(* IEC 61131-3 sources: plcassist-cli/packages/volt-lsp-iec/test-corpus/awa-palletizer/Device/Plc Logic/Application/Library Manager/AlarmManager (part 3) *)

(* ---- DATABASEFILEALARMSTORAGE.fb ---- *)
FUNCTION_BLOCK DATABASEFILEALARMSTORAGE EXTENDS AlarmStorageManager
VAR
	M_SAPPLICATIONNAME : STRING;
	M_AITFALARMSTORAGELISTENER : ARRAY [0..(COUNT_MAX_ALARM_STORAGE_LISTENER - 1)] OF IAlarmStorageListener;
	M_SOLDREMOTEDEVICENAME : STRING;
	M_LIREMOTEDEVICENAMEVALUE : LINT;
	M_CACHEDDBVERSION : INT := UNDETERMINED_DB_VERSION;
	M_CACHEDDBVERSIONERROR : STO.ERROR;
	M_WRITECONTEXT : DatabaseFileWriteContext;
	M_XCHANGESTATETONORMAL : BOOL;
	M_XASSIGNINACTIVETIMESTAMPS : BOOL;
	COUNT_MAX_ALARM_STORAGE_LISTENER : INT := 5;
	UNDETERMINED_DB_VERSION : INT := -1;
	ASSIGNINACTIVETIMESTAMPS : BOOL;
	CHANGESTATETONORMAL : BOOL;
	TABLE : STO.ITable;
	WRITEACCESSNECESSARY : BOOL;
END_VAR
END_FUNCTION_BLOCK

METHOD GETDATABASEFILEPATH : STRING
END_METHOD

METHOD GETFILELIMIT : FileLimit
END_METHOD

METHOD GETMAXRECORDCOUNT : UDINT
END_METHOD

METHOD GETSUBDIRECTORY : STRING
END_METHOD

METHOD WRITETOSTORAGE : STO.ERROR
VAR_INPUT
	ITFTABLE : STO.ITable;
	ROW : AlarmStorageRow;
	ICOUNTRETRIES : INT;
END_VAR
END_METHOD

METHOD CLEARBUFFER
END_METHOD

METHOD ADDALARMSTORAGELISTENER : EAlarmStorageReaderErrors
VAR_INPUT
	ITFALARMSTORAGELISTENER : IAlarmStorageListener;
END_VAR
END_METHOD

METHOD CREATEALARMSTORAGEMETADATAFILE
VAR_INPUT
	UDICOUNTCOLUMNSTBLALARM : CAA.COUNT;
END_VAR
END_METHOD

METHOD OPENTABLE2 : STO.ITable
VAR_INPUT
	XREADONLY : BOOL;
END_VAR
VAR_OUTPUT
	EERROR : STO.ERROR;
END_VAR
END_METHOD

METHOD REMOVEALARMSTORAGELISTENER : EAlarmStorageReaderErrors
VAR_INPUT
	ITFALARMSTORAGELISTENER : IAlarmStorageListener;
END_VAR
END_METHOD

METHOD CHECKFILELIMITREACHED : STO.Error
VAR_INPUT
	ITFTABLE : STO.ITable;
	ICOUNTRETRIES : INT;
	ICOUNTROWSTOINSERT : INT;
END_VAR
END_METHOD

METHOD GETEXCLUSIVETRANSACTION : STO.ITransaction
VAR_INPUT
	ICOUNTRETRIES : INT;
END_VAR
VAR_OUTPUT
	EERROR : STO.ERROR;
END_VAR
END_METHOD

METHOD WRITETOSTORAGE2 : STO.ERROR
VAR_INPUT
	ITFTABLE : STO.ITable;
	ROW : AlarmStorageRow;
	ITFTRANSACTION : STO.ITransaction;
END_VAR
END_METHOD

METHOD DELETEALARMSTORAGEFILE : STO.ERROR
VAR_INPUT
	SFILEPATH : CAA.FILENAME;
END_VAR
END_METHOD

METHOD GETALARMSFROMSTORAGE : STO.ERROR
VAR_INPUT
	ISKIPROWS : INT;
	IMAXROWS : INT;
	FILTERCRITERIA : REFERENCE TO VisuFbAlarmFilterCriteria;
	ITFALARMDATABLOCK : IAlarmDataBlockBase2;
END_VAR
VAR_IN_OUT
	BROWIDVALID : BOOL;
	DIROWID : DINT;
END_VAR
END_METHOD

METHOD GETCOUNTALARMSFROMSTORAGE : DINT
VAR_INPUT
	FILTERCRITERIA : REFERENCE TO VisuFbAlarmFilterCriteria;
	ITFALARMDATABLOCK : IAlarmDataBlockBase2;
END_VAR
VAR_OUTPUT
	EERROR : STO.ERROR;
	DWCOUNTLATCHVARIABLESINSTORAGE : CAA.COUNT;
END_VAR
END_METHOD

METHOD CREATEWRITECONTEXT : IDatabaseFileWriteContext
END_METHOD

METHOD SCANSTORAGE : STO.ERROR
VAR_INPUT
	ITFCONSUMER : IRemoteDeviceTraversalConsumer;
END_VAR
VAR_OUTPUT
	IVERSION : INT;
	DIREMOTEENTRIESCNT : DINT;
END_VAR
END_METHOD

METHOD WRITETOSTORAGE3 : STO.ERROR
VAR_INPUT
	WRITECONTEXT : IDatabaseFileWriteContext;
	ROW : AlarmStorageRow;
	XFORCEINSERT : BOOL;
	XFIRST : BOOL;
END_VAR
END_METHOD

METHOD CLEARALARMSINSTATENORMAL : STO.Error
VAR_INPUT
	ITFTABLE : STO.ITable;
END_VAR
VAR_OUTPUT
	XFINISHED : BOOL;
END_VAR
VAR_IN_OUT
	DIREMAININGROWCOUNT : DINT;
END_VAR
END_METHOD

METHOD ROWSELECT : STO.IRow
VAR_INPUT
	ITFTABLE : STO.ITable;
	IDROW : CAA.IDENT;
END_VAR
END_METHOD

METHOD CHECKRECORDLIMITREACHED : STO.Error
VAR_INPUT
	ITFTABLE : STO.ITable;
	ICOUNTRETRIES : INT;
	ICOUNTROWSTOINSERT : INT;
	XFORCE : BOOL;
END_VAR
VAR_OUTPUT
	XLIMIT : BOOL;
	UDIMAXRECORDCOUNT : UDINT;
END_VAR
END_METHOD

METHOD DELETEALARMS : STO.Error
VAR_INPUT
	ITFTABLE : STO.ITable;
	ICOUNTRETRIES : INT;
	DICOUNTROWSTODELETE : DINT;
END_VAR
VAR_OUTPUT
	DIROWSDELETED : DINT;
END_VAR
END_METHOD

METHOD GETRECORDSIZE : INT
END_METHOD

METHOD GETSTORAGESIZE : LINT
END_METHOD

METHOD SETEMPTYTIMESTAMPINACTIVETOSTARTTIME : STO.Error
VAR_INPUT
	ITFTABLE : STO.ITable;
END_VAR
END_METHOD

METHOD CHECKFILELIMITREACHEDUDINT : STO.ERROR
VAR_INPUT
	ITFTABLE : STO.ITable;
	ICOUNTRETRIES : INT;
	UDICOUNTROWSTOINSERT : UDINT;
END_VAR
END_METHOD

METHOD CHECKRECORDLIMITREACHEDUDINT : STO.ERROR
VAR_INPUT
	ITFTABLE : STO.ITable;
	ICOUNTRETRIES : INT;
	UDICOUNTROWSTOINSERT : UDINT;
	XFORCE : BOOL;
END_VAR
VAR_OUTPUT
	XLIMIT : BOOL;
	UDIMAXRECORDCOUNT : UDINT;
END_VAR
END_METHOD

METHOD PRVCHECKFILELIMITREACHED : STO.Error
VAR_INPUT
	ITFTABLE : STO.ITable;
	ICOUNTRETRIES : INT;
	UDICOUNTROWSTOINSERT : UDINT;
END_VAR
END_METHOD

METHOD PRVCHECKRECORDLIMITREACHED : STO.Error
VAR_INPUT
	ITFTABLE : STO.ITable;
	ICOUNTRETRIES : INT;
	UDICOUNTROWSTOINSERT : UDINT;
	XFORCE : BOOL;
END_VAR
VAR_OUTPUT
	XLIMIT : BOOL;
	UDIMAXRECORDCOUNT : UDINT;
END_VAR
END_METHOD

METHOD PRVDELETEALARMSTOREACHLIMIT : BOOL
VAR_INPUT
	ITFTABLE : STO.ITable;
	ICOUNTRETRIES : INT;
	UDICOUNTROWSTODELETE : UDINT;
END_VAR
VAR_OUTPUT
	IROWSDELETED : INT;
	EERROR : STO.ERROR;
END_VAR
END_METHOD

METHOD PRVFINDLATCHVARSTRING
VAR_INPUT
	CBPINPUTSTRING : CharBufferPtr;
	BYTYPECLASS : BYTE;
	IVERSION : INT;
	ITFTABLE : STO.ITable;
END_VAR
VAR_OUTPUT
	DIROWID : DINT;
	XFOUND : BOOL;
END_VAR
VAR_IN_OUT
	EERROR : STO.ERROR;
	WSINPUTSTRING : WSTRING(255);
END_VAR
END_METHOD

METHOD PRVFINDLATCHVARSTRING_DBVERBEFORE5
VAR_INPUT
	CBPINPUTSTRING : CharBufferPtr;
	BYTYPECLASS : BYTE;
	ITFCURSOR : STO.ICursor;
END_VAR
VAR_OUTPUT
	DIROWID : DINT;
	XFOUND : BOOL;
END_VAR
VAR_IN_OUT
	EERROR : STO.ERROR;
END_VAR
END_METHOD

METHOD PRVFINDLATCHVARSTRING_DBVERRECENT
VAR_INPUT
	ITFCURSOR : STO.ICursor;
END_VAR
VAR_OUTPUT
	DIROWID : DINT;
	XFOUND : BOOL;
END_VAR
VAR_IN_OUT
	EERROR : STO.ERROR;
	WSINPUTSTRING : WSTRING(255);
END_VAR
END_METHOD

METHOD PRVGETDATABASEFILEPATH : STRING
VAR_INPUT
	SVERSIONINCOMPATIBLECHANGE : STRING;
END_VAR
VAR_OUTPUT
	EERROR : STO.ERROR;
END_VAR
END_METHOD

METHOD PRVGETVERSION : STO.ERROR
VAR_OUTPUT
	IVERSION : INT;
END_VAR
END_METHOD

METHOD PRVGETVERSIONFROMDATABASE : STO.ERROR
VAR_OUTPUT
	IVERSION : INT;
END_VAR
END_METHOD

METHOD PRVREMOVERECORDLIMITREACHED : STO.Error
VAR_INPUT
	UDIMAXRECORDCOUNT : UDINT;
	ITFTABLE : STO.ITable;
	ICOUNTRETRIES : INT;
	ICOUNTROWSTOINSERT : UDINT;
END_VAR
END_METHOD

METHOD PRVSEARCHMINROWIDS : STO.ERROR
VAR_INPUT
	ITFTABLE : STO.ITable;
	ICOUNTROWSIDSTOSEARCH : INT;
	PADWROWIDS : POINTER TO ARRAY [0..50] OF CAA.IDENT;
	IEFFECTIVEARRAYSIZE : INT;
END_VAR
VAR_OUTPUT
	ICOUNTROWSIDS : INT;
END_VAR
END_METHOD

METHOD PRVSETTYPEDVALUE : STO.ERROR
VAR_INPUT
	BYTYPECLASS : BYTE;
	LIVALUE : LINT;
	ITFROWBASE : STO.IRowBase;
	COLVALUE : CAA.IDENT;
	COLTYPE : CAA.IDENT;
END_VAR
END_METHOD

METHOD PRVSORTROWIDS
VAR_INPUT
	PADWROWIDS : POINTER TO ARRAY [0..0] OF CAA.IDENT;
	NFIRST : INT;
	NLAST : INT;
END_VAR
END_METHOD

METHOD PRVSTOREALARMCOMMENTS : STO.ERROR
VAR_INPUT
	PROW : POINTER TO AlarmStorageRow;
	ITFROWPLANCHET : STO.IRowPlanchet;
	ITFROW : STO.IRow;
END_VAR
END_METHOD

METHOD PRVUPDATEROW : BOOL
VAR_INPUT
	HTASK : RTS_IEC_HANDLE;
	ITFROW : STO.IRow;
	ICOUNTRETRIES : INT;
	EERROR : STO.ERROR;
END_VAR
END_METHOD

METHOD PRVWRITEALARMCOMMENTCOLUMN
VAR_INPUT
	PWSVALUE : POINTER TO WSTRING;
	ITFROWPLANCHET : STO.IRowPlanchet;
	ITFROW : STO.IRow;
	DATABASEIDENT : CAA.IDENT;
	ERRACTION : INT;
END_VAR
VAR_IN_OUT
	EERROR : STO.ERROR;
END_VAR
END_METHOD

METHOD PRVWRITEBYTEORDERFLAG
END_METHOD

METHOD PRVWRITELATCHVARSTRINGS
VAR_INPUT
	ITFROWBASE : STO.IRowBase;
	PROW : POINTER TO AlarmStorageRow;
	WRITECONTEXT : IDatabaseFileWriteContext;
END_VAR
VAR_IN_OUT
	EERROR : STO.ERROR;
END_VAR
END_METHOD

METHOD PRVWRITETOSTORAGE : STO.ERROR
VAR_INPUT
	WRITECONTEXT : IDatabaseFileWriteContext;
	ROW : AlarmStorageRow;
	ICOUNTRETRIES : INT;
	XCHECKFILELIMITREACHED : BOOL;
	XFORCEINSERT : BOOL;
END_VAR
END_METHOD

METHOD PRVWRITETOTBLLATCHVARSTRINGS : STO.ERROR
VAR_INPUT
	WRITECONTEXT : IDatabaseFileWriteContext;
	CBPINPUTSTRING : CharBufferPtr;
	BYTYPECLASS : BYTE;
END_VAR
VAR_OUTPUT
	DIROWID : DINT;
END_VAR
END_METHOD

METHOD PRVWRITETRIGGERVALUE
VAR_INPUT
	ITFROWBASE : STO.IRowBase;
	BYTRIGGERVALUETYPE : BYTE;
	LITRIGGERVALUEVAL : LINT;
END_VAR
VAR_IN_OUT
	EERROR : STO.ERROR;
END_VAR
END_METHOD

(* ---- DATABASEFILEWRITECONTEXT.fb ---- *)
FUNCTION_BLOCK DATABASEFILEWRITECONTEXT EXTENDS DatabaseFileWriteContextBase
VAR
	_INUSE : BOOL;
	M_ICOUNTRETRIES : INT := AlarmConstants.RETRY_COUNT;
	M_ICOUNTCYCLEWAIT : INT;
END_VAR
END_FUNCTION_BLOCK

METHOD INITIALIZE : BOOL
VAR_IN_OUT
	DB : DatabaseFileAlarmStorage;
END_VAR
END_METHOD

METHOD RELEASE
VAR_INPUT
	EERRORFORCOMMIT : STO.ERROR;
END_VAR
END_METHOD

METHOD PRVINCREASERETRYCOUNT : BOOL
END_METHOD

METHOD PRVRESETRETRYCOUNT : BOOL
END_METHOD

(* ---- DATABASEFILEWRITECONTEXTBASE.fb ---- *)
FUNCTION_BLOCK DATABASEFILEWRITECONTEXTBASE
VAR
	_MAINTABLE : STO.ITable;
	_STRINGLATCHTABLE : STO.ITable;
	_TRANSACTION : STO.ITransaction;
	_STORAGEMAN : REFERENCE TO DatabaseFileAlarmStorage;
	MAINTABLE : STO.ITable;
	TRANSACTION : STO.ITransaction;
END_VAR
END_FUNCTION_BLOCK

METHOD GETSTRINGLATCHTABLE : STO.ITable
VAR_OUTPUT
	EERROR : STO.ERROR;
END_VAR
END_METHOD

METHOD RELEASE
VAR_INPUT
	EERRORFORCOMMIT : STO.ERROR;
END_VAR
END_METHOD

(* ---- DATABASEFILEWRITECONTEXTTEMPORARY.fb ---- *)
FUNCTION_BLOCK DATABASEFILEWRITECONTEXTTEMPORARY EXTENDS DatabaseFileWriteContextBase
END_FUNCTION_BLOCK

METHOD FB_EXIT : BOOL
VAR_INPUT
	BINCOPYCODE : BOOL;
END_VAR
END_METHOD

METHOD INITIALIZE : BOOL
VAR_INPUT
	MAINTABLE : STO.ITable;
	TRANSACTION : STO.ITransaction;
END_VAR
VAR_IN_OUT
	STORAGEMAN : DatabaseFileAlarmStorage;
END_VAR
END_METHOD

(* ---- DATABASESIZELIMIT.fb ---- *)
FUNCTION_BLOCK DATABASESIZELIMIT
VAR
	M_XINITIALIZED : BOOL;
	M_XFIRST : BOOL := TRUE;
	M_XFIRSTREMOVE : BOOL := TRUE;
	M_METRICS : STO.METRICS;
	M_ITFDATABASEFILEALARMSTORAGE7 : IDatabaseFileAlarmStorage7;
	M_ITFALARMSTORAGEMANAGER : IAlarmStorageManager;
	M_SYSRECORDSIZE : INT;
	M_LISTORAGESIZE : LINT;
	M_XERRORDISPLAYED : BOOL;
	M_LIFILESIZEINERROR : LINT;
	M_ICNTREORGERR : INT;
	M_XBLOCKED : BOOL;
	M_ITEMPREDUCTIONRECORDNUM : INT;
	M_TLASTREORGTIME : TIME;
	M_ICNTDBREORD : INT;
	ISBLOCKED : BOOL;
	LASTREORDERINGTIME : TIME;
	REORDERINGCOUNT : INT;
END_VAR
END_FUNCTION_BLOCK

METHOD CHECKFORSIZELIMIT : BOOL
END_METHOD

METHOD INITIALIZE
VAR_INPUT
	ITFDATABASEFILEALARMSTORAGE : IDatabaseFileAlarmStorage;
END_VAR
END_METHOD

METHOD PRVDBMETRICS : STO.ERROR
VAR_OUTPUT
	MMETRICS : STO.METRICS;
END_VAR
END_METHOD

METHOD PRVGETRECORDSIZE : INT
END_METHOD

METHOD PRVGETRECORDSTOREMOVE : DINT
VAR_INPUT
	LIBYTESTOREMOVE : LINT;
END_VAR
VAR_OUTPUT
	IRECORDSIZE : INT;
END_VAR
END_METHOD

METHOD PRVREORGDB : STO.ERROR
END_METHOD

(* ---- DEFAULTALARMFILTERCRITERIA.fb ---- *)
FUNCTION_BLOCK DEFAULTALARMFILTERCRITERIA
END_FUNCTION_BLOCK

METHOD AREALLALARMCLASSESSELECTED : BOOL
END_METHOD

METHOD AREALLALARMGROUPSSELECTED : BOOL
END_METHOD

METHOD GETALARMCLASSES : POINTER TO ARRAY [0..0] OF UDINT
END_METHOD

METHOD GETALARMGROUPS : POINTER TO ARRAY [0..0] OF UDINT
END_METHOD

METHOD GETCOUNTALARMCLASSES : INT
END_METHOD

METHOD GETCOUNTALARMGROUPS : INT
END_METHOD

METHOD GETPRIORITYFROM : USINT
END_METHOD

METHOD GETPRIORITYTO : USINT
END_METHOD

(* ---- EVENTDISPATCHER.fb ---- *)
FUNCTION_BLOCK EVENTDISPATCHER
VAR
	_HGETCOUNTEVENT : RTS_IEC_HANDLE := Events.Invalid_Handle;
	_HGETCOUNTEVENTINTERFACE : RTS_IEC_HANDLE := Events.Invalid_Handle;
	_HGETALARMSEVENT : RTS_IEC_HANDLE := Events.Invalid_Handle;
	_HGETALARMSEVENTINTERFACE : RTS_IEC_HANDLE := Events.Invalid_Handle;
	_HCHANNELCLOSEDEVENT : RTS_IEC_HANDLE := Events.Invalid_Handle;
	_HCHANNELCLOSEDEVENTINTERFACE : RTS_IEC_HANDLE := Events.Invalid_Handle;
	_HHANDLESERVICEEVENT : RTS_IEC_HANDLE := Events.Invalid_Handle;
	_HHANDLESERVICEEVENTINTERFACE : RTS_IEC_HANDLE := Events.Invalid_Handle;
	_SERVICEHANDLER : AlarmServiceHandler;
END_VAR
END_FUNCTION_BLOCK

METHOD EVENTCALLBACK : UDINT
VAR_INPUT
	PEVENTPARAM : POINTER TO EventParam;
END_VAR
END_METHOD

METHOD FB_EXIT : BOOL
VAR_INPUT
	BINCOPYCODE : BOOL;
END_VAR
END_METHOD

METHOD FB_INIT : BOOL
VAR_INPUT
	BINITRETAINS : BOOL;
	BINCOPYCODE : BOOL;
END_VAR
END_METHOD

(* ---- EXPRESSIONOBSERVATIONTYPE.fb ---- *)
FUNCTION_BLOCK EXPRESSIONOBSERVATIONTYPE
VAR_INPUT
	M_UIID : ALARM_ID;
	M_EXPRESSIONEVALUATOR : IExpressionEvaluator;
END_VAR
END_FUNCTION_BLOCK

METHOD ISACTIVE : BOOL
VAR_INPUT
	ECURRSTATE : AlarmState;
END_VAR
END_METHOD

METHOD ISIMMEDIATELYACTIVE : BOOL
END_METHOD

(* ---- FORMATSTRINGSCANNER.fb ---- *)
FUNCTION_BLOCK FORMATSTRINGSCANNER
END_FUNCTION_BLOCK

METHOD GETFORMATSTRING : BOOL
VAR_INPUT
	RCBSMESSAGE : REFERENCE TO CharBufferString;
	PCBSPLACEHOLDER : POINTER TO CharBufferString;
	IOFFSET : INT;
	ILENGTHPREFIX : INT;
END_VAR
VAR_OUTPUT
	SFORMATSTRING : STRING;
	ITOTALPLACEHOLDERLENGTH : INT;
END_VAR
END_METHOD

(* ---- HASHTABLEKEYELEMENT.fb ---- *)
FUNCTION_BLOCK HASHTABLEKEYELEMENT EXTENDS InstanceBase
VAR
	_INSTANCEPOINTER : POINTER TO BYTE;
	_ALARMTEMPLATENAME : POINTER TO STRING;
	_LIHASH : LINT;
	ALARMTEMPLATENAME : POINTER TO STRING;
	INSTANCEPOINTER : POINTER TO BYTE;
END_VAR
END_FUNCTION_BLOCK

METHOD ELEMENTCOMPARETO : INT
VAR_INPUT
	ITFELEMENT : COL.IElement;
END_VAR
END_METHOD

METHOD ELEMENTEQUALS : BOOL
VAR_INPUT
	ITFELEMENT : COL.IElement;
END_VAR
END_METHOD

METHOD ELEMENTHASHCODE : LINT
END_METHOD

METHOD PRVCALCULATEHASH : LINT
END_METHOD

METHOD PRVINSTINIT : COL.FBF.ERROR
VAR_INPUT
	ITFDATA : COL.FBF.IData;
END_VAR
END_METHOD

(* ---- HASHTABLEKEYELEMENTDATA.fb ---- *)
FUNCTION_BLOCK HASHTABLEKEYELEMENTDATA EXTENDS InstanceData
VAR_INPUT
	PALARMINSTANCE : POINTER TO BYTE;
	STALARMTEMPLATENAME : POINTER TO STRING;
END_VAR
END_FUNCTION_BLOCK

(* ---- HASHTABLEKEYELEMENTFACTORY.fb ---- *)
FUNCTION_BLOCK HASHTABLEKEYELEMENTFACTORY EXTENDS FactoryBase
VAR
	PRVINSTCOUNT : CAA.COUNT;
	PRVINSTPOOLEXTENDSFACTOR : USINT;
	PRVINSTSIZE : CAA.SIZE;
END_VAR
END_FUNCTION_BLOCK

METHOD CREATE : IHashtableKeyElement
VAR_INPUT
	INSTANCEPOINTER : POINTER TO BYTE;
	PSTALARMTEMPLATENAME : POINTER TO STRING;
END_VAR
VAR_OUTPUT
	EERROR : COL.FBF.ERROR;
END_VAR
END_METHOD

(* ---- HASHTABLEVALUEELEMENT.fb ---- *)
FUNCTION_BLOCK HASHTABLEVALUEELEMENT EXTENDS InstanceBase
VAR
	_UDIALARMGROUPID : UDINT;
	_UITEMPLATEALARMSOFFSET : UINT;
	_UITEMPLATEALARMSLENGTH : UINT;
	_UITEMPLATEEVENTSOFFSET : UINT;
	_UITEMPLATEEVENTSLENGTH : UINT;
	ALARMGROUPID : UDINT;
	TEMPLATEALARMSLENGTH : UINT;
	TEMPLATEALARMSOFFSET : UINT;
	TEMPLATEEVENTSLENGTH : UINT;
	TEMPLATEEVENTSOFFSET : UINT;
END_VAR
END_FUNCTION_BLOCK

METHOD ELEMENTCOMPARETO : INT
VAR_INPUT
	ITFELEMENT : COL.IElement;
END_VAR
END_METHOD

METHOD ELEMENTEQUALS : BOOL
VAR_INPUT
	ITFELEMENT : COL.IElement;
END_VAR
END_METHOD

METHOD ELEMENTHASHCODE : LINT
END_METHOD

METHOD PRVINSTINIT : COL.FBF.ERROR
VAR_INPUT
	ITFDATA : COL.FBF.IData;
END_VAR
END_METHOD

(* ---- HASHTABLEVALUEELEMENTDATA.fb ---- *)
FUNCTION_BLOCK HASHTABLEVALUEELEMENTDATA EXTENDS InstanceData
VAR_INPUT
	UDIALARMGROUPID : UDINT;
	UITEMPLATEALARMSOFFSET : UINT;
	UITEMPLATEALARMSLENGTH : UINT;
	UITEMPLATEEVENTSOFFSET : UINT;
	UITEMPLATEEVENTSLENGTH : UINT;
END_VAR
END_FUNCTION_BLOCK

(* ---- HASHTABLEVALUEELEMENTFACTORY.fb ---- *)
FUNCTION_BLOCK HASHTABLEVALUEELEMENTFACTORY EXTENDS FactoryBase
VAR
	PRVINSTCOUNT : CAA.COUNT;
	PRVINSTPOOLEXTENDSFACTOR : USINT;
	PRVINSTSIZE : CAA.SIZE;
END_VAR
END_FUNCTION_BLOCK

METHOD CREATE : IHashtableValueElement
VAR_INPUT
	UDIALARMGROUPID : UDINT;
	UITEMPLATEALARMSOFFSET : UINT;
	UITEMPLATEALARMSLENGTH : UINT;
	UITEMPLATEEVENTSOFFSET : UINT;
	UITEMPLATEEVENTSLENGTH : UINT;
END_VAR
VAR_OUTPUT
	EERROR : COL.FBF.ERROR;
END_VAR
END_METHOD

(* ---- HISTORICALALARMMOCK.fb ---- *)
FUNCTION_BLOCK HISTORICALALARMMOCK EXTENDS ProxyFbAlarmHistorical
VAR_INPUT
	M_BALARMSTORAGE : BYTE;
	M_DWROWIDFIRST : DWORD;
	M_DWROWIDLAST : DWORD;
	M_SVALUE : STRING;
	M_WSVALUE : WSTRING;
END_VAR
END_FUNCTION_BLOCK

METHOD SETVALUES
VAR_INPUT
	ISET : INT;
END_VAR
END_METHOD

(* ---- LISTELEMENT.fb ---- *)
FUNCTION_BLOCK LISTELEMENT EXTENDS InstanceBase
VAR
	_ALARMINST : Alarm;
	_USICOUNTLATCHVARIABLES : USINT;
	_ARRLATCHVARIABLES : ARRAY [0..255] OF ValueTypeBundle;
	_XISACTIVEALARM : BOOL;
	ALARM : POINTER TO Alarm;
	ISACTIVEALARM : BOOL;
	ISDEACTIVATEDPREV : BOOL;
END_VAR
END_FUNCTION_BLOCK

METHOD ELEMENTCOMPARETO : INT
VAR_INPUT
	ITFELEMENT : COL.IElement;
END_VAR
END_METHOD

METHOD ELEMENTEQUALS : BOOL
VAR_INPUT
	ITFELEMENT : COL.IElement;
END_VAR
END_METHOD

METHOD ELEMENTHASHCODE : LINT
END_METHOD

METHOD GETLATCHVARIABLES : BOOL
VAR_OUTPUT
	PALATCHVARIABLES : POINTER TO ARRAY [0..255] OF ValueTypeBundle;
	USICOUNTLATCHVARIABLES : USINT;
END_VAR
END_METHOD

METHOD SETLATCHVARIABLES : BOOL
VAR_INPUT
	PALARM : POINTER TO Alarm;
END_VAR
END_METHOD

METHOD PRVINSTINIT : COL.FBF.ERROR
VAR_INPUT
	ITFDATA : COL.FBF.IData;
END_VAR
END_METHOD

(* ---- LISTELEMENTDATA.fb ---- *)
FUNCTION_BLOCK LISTELEMENTDATA EXTENDS InstanceData
END_FUNCTION_BLOCK

(* ---- LISTELEMENTFACTORY.fb ---- *)
FUNCTION_BLOCK LISTELEMENTFACTORY EXTENDS FactoryBase
VAR
	PRVINSTCOUNT : CAA.COUNT;
	PRVINSTPOOLEXTENDSFACTOR : USINT;
	PRVINSTSIZE : CAA.SIZE;
END_VAR
END_FUNCTION_BLOCK

METHOD CREATE : IListElement
VAR_OUTPUT
	EERROR : COL.FBF.ERROR;
END_VAR
END_METHOD

(* ---- MESSAGECOMPARER.fb ---- *)
FUNCTION_BLOCK MESSAGECOMPARER EXTENDS TSLastComparer
VAR
	M_STRINGTYPE : __SYSTEM.TYPE_CLASS;
	M_IWHICHMESSAGE : INT;
	M_ICOUNTLATCHVARIABLES : INT;
	M_CBSMESSAGE1 : CharBufferString;
	M_CBSMESSAGE2 : CharBufferString;
	M_CBSMESSAGE1REPLACED : CharBufferString;
	M_CBSMESSAGE2REPLACED : CharBufferString;
	M_ABYBUFFERMESSAGE1REPLACED : ARRAY [0..(BUFFER_LENGTH - 1)] OF BYTE;
	M_ABYBUFFERMESSAGE2REPLACED : ARRAY [0..(BUFFER_LENGTH - 1)] OF BYTE;
	M_TIMESTAMPANDVALUESCONTAINER : TimestampAndValuesContainer;
	BUFFER_LENGTH : INT := (2 * (255 + 1));
END_VAR
END_FUNCTION_BLOCK

METHOD BEFORECOMPARE
VAR_INPUT
	STRINGTYPE : __SYSTEM.TYPE_CLASS;
	IWHICHMESSAGE : INT;
	ICOUNTLATCHVARIABLES : INT;
END_VAR
END_METHOD

METHOD COMPARE : INT
VAR_INPUT
	DIINDEXALARM1 : DINT;
	DIINDEXALARM2 : DINT;
END_VAR
END_METHOD

METHOD PRVGETALARMMESSAGE : CharBufferPtr
VAR_INPUT
	UDIALARMGROUPID : UDINT;
	UDIALARMID : UDINT;
	SDEVICENAME : STRING;
END_VAR
VAR_OUTPUT
	SALARMID : STRING;
END_VAR
END_METHOD

METHOD PRVREPLACEPLACEHOLDERS : BOOL
VAR_INPUT
	DIINDEXALARM : DINT;
	CBPMESSAGE : CharBufferPtr;
	RCBSMESSAGE : REFERENCE TO CharBufferString;
	RCBSMESSAGEREPLACED : REFERENCE TO CharBufferString;
END_VAR
END_METHOD

(* ---- ONLYDATEANDTIMEPLACEHOLDER.fb ---- *)
FUNCTION_BLOCK ONLYDATEANDTIMEPLACEHOLDER
VAR
	M_APLACEHOLDEROCCURRENCE : ARRAY [PLACEHOLDER_DATE..PLACEHOLDER_TIME] OF PlaceholderOccurrence;
	PLACEHOLDER_DATE : INT := 0;
	PLACEHOLDER_TIME : INT := 1;
END_VAR
END_FUNCTION_BLOCK

METHOD FB_INIT : BOOL
VAR_INPUT
	BINITRETAINS : BOOL;
	BINCOPYCODE : BOOL;
END_VAR
END_METHOD

METHOD ANALYZEPLACEHOLDERS
VAR_INPUT
	STRINGTYPE : __SYSTEM.TYPE_CLASS;
END_VAR
END_METHOD

METHOD GETCOUNTPLACEHOLDERS : SINT
END_METHOD

METHOD GETPLACEHOLDER : PlaceholderOccurrence
VAR_INPUT
	SIWHICHPLACEHOLDER : SINT;
END_VAR
END_METHOD

METHOD HASPLACEHOLDERREQUIRINGCYCLICALLYUPDATE : BOOL
END_METHOD

METHOD HASPLACEHOLDERS : BOOL
END_METHOD

METHOD ISOPTIMIZEDPLACEHOLDERREPLACEMENTSUPPORTED : BOOL
END_METHOD

(* ---- PRIORITYCOMPARER.fb ---- *)
FUNCTION_BLOCK PRIORITYCOMPARER EXTENDS TSLastComparer
END_FUNCTION_BLOCK

METHOD COMPARE : INT
VAR_INPUT
	DIINDEXALARM1 : DINT;
	DIINDEXALARM2 : DINT;
END_VAR
END_METHOD

(* ---- PROXY.fb ---- *)
FUNCTION_BLOCK PROXY
VAR
	M_XISINIT : BOOL;
	M_IRUNSTATUS : INT;
	M_ITFCOMMCHANNEL : IProxyCommChannel;
	M_ITEST : INT;
	M_ESTATE : ProxyEnumState;
	M_SDEVICENAME : STRING;
	M_LIBVERALMMAN : VERSION;
	M_LTSTARTTIMECHANNEL : LTIME;
	M_LTSTARTTIMERUN : LTIME;
	M_LTSTARTTIME : LTIME;
	M_ISTATE : INT;
	M_XALREADYDISP : BOOL;
	M_TTIMEOUT : TIME;
	M_IREQIDSENT : INT;
	M_IREQIDREC : INT;
	M_XWITHERRORS : BOOL;
	M_DWBASETIME : DWORD := (50 * 1000);
	M_DWACTALMTIME : DWORD := (200 * 1000);
	M_DWHISALMTIME : DWORD := (1000 * 1000);
	M_DWACKALMTIME : DWORD := (1000 * 1000);
	M_TGENTIMEOUT : TIME := DEFAULT_TIMEOUT;
	M_APROXYRUNTASKCALL : ARRAY [1..ProxyConstants.MAX_TASK] OF ProxyStructTaskCall;
	M_IRUNTASKCALLMAX : INT;
	M_APROXYPRERUNTASKCALL : ARRAY [1..ProxyConstants.MAX_TASK] OF ProxyStructTaskCall;
	M_IPRERUNTASKCALLMAX : INT;
	M_ITASKCALL : INT;
	M_SPROXYNAME : STRING;
	M_PSAPPNAME : POINTER TO STRING;
	M_CBSMESSAGE : CharBufferString;
	M_AWLOCALBUFFER : ARRAY [0..(LOCAL_TEXT_BUFFER_LENGTH / 2)] OF WORD;
	M_ARECORDS : ARRAY [0..(MAX_RECORDS - 1)] OF ProxyStructRecord;
	M_IRECINUSE : INT;
	M_SIHASSTORAGE : SINT := -1;
	M_DWROWIDFIRSTREMDB : DWORD := AlarmConstants.INVALID_ROWID;
	M_DWROWIDLASTREMDB : DWORD := AlarmConstants.INVALID_ROWID;
	M_DWROWIDLASTVALIDREAD : DWORD := AlarmConstants.INVALID_ROWID;
	M_DWROWIDLASTLOCDB : DWORD := AlarmConstants.INVALID_ROWID;
	M_IROWCOUNTTOREAD : INT;
	M_PAHISTALARMGROUPS : ARRAY [1..MAX_HIST_GROUPS] OF POINTER TO STRING;
	M_IHISTALARMGROUPSNUM : INT;
	M_IHISTRECORDID : INT := -1;
	M_XFIRSTHISTREADDONE : BOOL;
	M_XFIRSTHISTACTIVEREADDONE : BOOL;
	M_XDISP1DONE : BOOL;
	M_XDISP2DONE : BOOL;
	M_XDISP3DONE : BOOL;
	M_XDISP4DONE : BOOL;
	M_DIHISTACTIVEFIRSTENTRY : DINT;
	M_HISTACTIVEALMPENDINGQUEUE : ProxyFbHistActiveAlarmsQueue;
	M_HISTALMROWQUEUE : ProxyFbHistAlarmsRowQueue;
	M_HISTACTIVEALMROWQUEUE : ProxyFbHistAlarmsRowQueue;
	M_IHISTROWCOUNTREAD : INT;
	M_IHISTACTIVEROWCOUNTREAD : INT;
	M_TWRITEDBDURATIONTIME : TIME;
	M_IWRITEDBCNT : INT;
	M_DIWRITEDBCNTTOT : DINT;
	M_DISTORAGEROWSCOUNT : DINT;
	M_ISTORAGECLEAR : INT;
	M_ISTORAGECLEAROLD : INT := -1;
	M_IRECIXALMTOACK : INT;
	M_DIALMIXALMTOACK : DINT;
	M_LITIMELASTLOCDB : LINT;
	M_IVERSIONDB : INT;
	M_XCLIENTISREG : BOOL;
	M_HLOCKREADALM2 : RTS_IEC_HANDLE := RTS_INVALID_HANDLE;
	M_ICNTFORSTATISTICS : INT;
	M_DISTATHISTACTIVEALMSCNT : DINT;
	M_ISTATHISTROWALMSCNT : INT;
	M_ISTATHISTROWACTIVEALMSCNT : INT;
	_IRECORDID : INT;
	_DIALARMNUM : DINT;
	_ILATCHVARSNUM : INT;
	_IALARMCLASSNUM : INT;
	_XRAISEDMOREALARMSTHANSTORAGELIMITREPORTED : BOOL;
	STATE_IDLE : INT := 0;
	STATE_ANS_WAIT : INT := 10;
	RUN_START : INT := 0;
	RUN_RECORD : INT := 1;
	RUN_RECORD_HIST : INT := 2;
	RUN_PRERUN : INT := 3;
	RUN_CHECK_DATA : INT := 4;
	RUN_RUN : INT := 5;
	MAX_RECORDS : INT := 1;
	MAX_HIST_GROUPS : INT := 50;
	DEFAULT_NAME : STRING := '-Proxy-';
	DEFAULT_TIMEOUT : TIME := TIME#30s0ms;
	LOCAL_TEXT_BUFFER_LENGTH : INT := (1000 * 2);
	ACTIVEALARMSCOUNT : DINT;
	APPLICATION : POINTER TO STRING;
	HASSTORAGE : BOOL;
	HISTACTIVEALARMREAD : INT;
	HISTALARMREAD : INT;
	ISINITIALIZED : BOOL;
	ISRUNCYCLICOK : BOOL;
	LATCHVARSNUM : INT;
	MAXHISTROWSTOREAD : INT;
	PROXYTASKCALL : ARRAY [1..ProxyConstants.MAX_TASK] OF ProxyStructTaskCall;
	PROXYTASKCALLSIZE : INT;
	RECORDID : INT;
	RECORDIDHISTORICAL : INT;
	ROWIDFIRST : DWORD;
	ROWIDLAST : DWORD;
	ROWIDLASTREAD : DWORD;
	TOTALARMNUM : DINT;
	TOTCLASSNUM : INT;
END_VAR
END_FUNCTION_BLOCK

METHOD FB_EXIT : BOOL
VAR_INPUT
	BINCOPYCODE : BOOL;
END_VAR
END_METHOD

METHOD FB_INIT : BOOL
VAR_INPUT
	BINITRETAINS : BOOL;
	BINCOPYCODE : BOOL;
END_VAR
END_METHOD

METHOD CYCLICCALL : BOOL
END_METHOD

METHOD GETACTIVEALARMS : INT
VAR_INPUT
	SNAME : STRING;
	FILTERCRITERIA : REFERENCE TO VisuFbAlarmFilterCriteria;
	ITFALARMDATABLOCK : IAlarmDataBlockBaseDINT;
END_VAR
VAR_IN_OUT
	DISTUBPROG : DINT;
END_VAR
END_METHOD

METHOD GETACTIVEALARMS2
VAR_INPUT
	FILTERCRITERIA : REFERENCE TO VisuFbAlarmFilterCriteria;
	PAITFALARMS : POINTER TO ARRAY [0..10] OF IAlarm;
	DIARRSIZE : DINT;
END_VAR
VAR_OUTPUT
	DICOUNT : DINT;
END_VAR
END_METHOD

METHOD GETALARMCLASSDESC
VAR_INPUT
	UDIID : UDINT;
END_VAR
VAR_OUTPUT
	SDESC : ProxyStructAlarmClassDesc;
END_VAR
END_METHOD

METHOD GETALARMCLASSDESCBYNAME
VAR_INPUT
	SCLASSNAME : STRING;
END_VAR
VAR_OUTPUT
	SDESC : ProxyStructAlarmClassDesc;
END_VAR
END_METHOD

METHOD GETALARMDESC
VAR_INPUT
	UDIALMID : UDINT;
	UDIGRPID : UDINT;
END_VAR
VAR_OUTPUT
	SDESC : ProxyStructAlarmDesc;
END_VAR
END_METHOD

METHOD GETALARMDISPLAYOPTIONS
VAR_INPUT
	ITFALARMMETAOBJECTSTUB5 : IAlarmMetaObjectStub5;
	REFDISPLAYOPTIONS : REFERENCE TO DisplayOptions;
END_VAR
VAR_OUTPUT
	XVALID : BOOL;
	SCLASSREMAP : STRING;
END_VAR
END_METHOD

METHOD GETALARMGROUPDESC
VAR_INPUT
	UDIID : UDINT;
END_VAR
VAR_OUTPUT
	SDESC : ProxyStructAlarmGroupDesc;
END_VAR
END_METHOD

METHOD GETALARMGROUPDESCBYNAME
VAR_INPUT
	SGRPNAME : STRING;
END_VAR
VAR_OUTPUT
	SDESC : ProxyStructAlarmGroupDesc;
END_VAR
END_METHOD

METHOD GETALARMMESSAGE
VAR_INPUT
	ITFALARMMETAOBJECTSTUB5 : IAlarmMetaObjectStub5;
	IWHICHMESSAGE : INT;
	REFCHARBUFFERSTRING : REFERENCE TO CharBufferString;
	STRINGTYPE : __SYSTEM.TYPE_CLASS;
END_VAR
END_METHOD

METHOD GETALARMMESSAGE2 : Stu.CharBufferPtr
VAR_INPUT
	STEXTLISTNAME : STRING;
	STEXTLISTINDEX : STRING;
	IWHICHMESSAGE : INT;
	STRINGTYPE : __SYSTEM.TYPE_CLASS;
END_VAR
END_METHOD

METHOD GETPROXYNAME : POINTER TO STRING
END_METHOD

METHOD GETTOTALALARMSCOUNT : DINT
END_METHOD

METHOD INITIALIZE : BOOL
VAR_INPUT
	PPARAM : POINTER TO ProxyStructInitialize;
	ITEST : INT;
END_VAR
END_METHOD

METHOD REGISTERUSERCLIENT
END_METHOD

METHOD SETALARMSTOACK
VAR_INPUT
	ITFALARMMETAOBJECTSTUB : IAlarmMetaObjectStub5;
END_VAR
END_METHOD

METHOD SETINITIALDATAFROMDB
VAR_INPUT
	ROW : REFERENCE TO AlarmStorageRow;
	XFIRST : BOOL;
	IVERSION : INT;
END_VAR
END_METHOD

METHOD SETPARAMS
VAR_INPUT
	PPARAM : POINTER TO ProxyStructParam;
END_VAR
END_METHOD

METHOD COMMUNICATIONFINISHED
VAR_INPUT
	IREQUESTID : INT;
	XWITHERRORS : BOOL;
END_VAR
END_METHOD

METHOD PROXYMANAGERLOG
VAR_INPUT
	SVAL1 : STRING(255);
	SVAL2 : STRING(255);
	SVAL3 : STRING(255);
	UDISEV : UDINT;
END_VAR
END_METHOD

METHOD SETACTIVEALARMSCOUNT
VAR_INPUT
	DICOUNT : DINT;
END_VAR
END_METHOD

METHOD SETALARMMANAGERLIBVERSION
VAR_INPUT
	LIBVER : VERSION;
END_VAR
END_METHOD

METHOD SETDEVICENAME
VAR_INPUT
	SNAME : STRING;
END_VAR
END_METHOD

METHOD SETHASSTORAGE
VAR_INPUT
	XVALUE : BOOL;
END_VAR
END_METHOD

METHOD SETHISTACTIVEALARMSREAD
VAR_INPUT
	ICOUNT : INT;
END_VAR
END_METHOD

METHOD SETHISTALARMSREAD
VAR_INPUT
	DWROWIDLAST : DWORD;
	ICOUNT : INT;
	DISTORAGEROWSCOUNT : DINT;
	ISTORAGECLEAR : INT;
END_VAR
END_METHOD

METHOD SETLATCHVARSCOUNT
VAR_INPUT
	ICOUNT : INT;
END_VAR
END_METHOD

METHOD SETRECORDID
VAR_INPUT
	IVALUE : INT;
END_VAR
END_METHOD

METHOD SETROWIDS
VAR_INPUT
	DWROWIDFIRST : DWORD;
	DWROWIDLAST : DWORD;
END_VAR
END_METHOD

METHOD SETTOTALALARMSCOUNT
VAR_INPUT
	DICOUNT : DINT;
END_VAR
END_METHOD

METHOD SETTOTALCLASSESCOUNT
VAR_INPUT
	ICOUNT : INT;
END_VAR
END_METHOD

METHOD GETALARMGROUP : STRING
VAR_INPUT
	IWHICHALARMGROUP : INT;
END_VAR
END_METHOD

METHOD GETALARMGROUPSNUM : INT
END_METHOD

METHOD GETAPPLICATION : STRING
END_METHOD

METHOD GETCOUNTALARMSTOACKNOWLEDGE : INT
END_METHOD

METHOD GETNEXTALARMTOACKNOWLEDGE : BOOL
VAR_INPUT
	XFISRTENTRY : BOOL;
END_VAR
VAR_OUTPUT
	ALARMTOACKNOWLEDGE : AlarmToAcknowledge;
END_VAR
END_METHOD

METHOD GETPROXYACTIVEALARMOBJECT : IProxyAlarmObject
VAR_INPUT
	DIOBJNUM : DINT;
END_VAR
END_METHOD

METHOD GETPROXYALARMCLASSDESCRIPTIONOBJECT : POINTER TO ProxyStructAlarmClass
VAR_INPUT
	IOBJNUM : INT;
END_VAR
END_METHOD

METHOD GETPROXYALARMDESCRIPTIONOBJECT : POINTER TO ProxyStructAlarm
VAR_INPUT
	IOBJNUM : INT;
END_VAR
END_METHOD

METHOD GETPROXYALARMGROUPDESCRIPTIONOBJECT : POINTER TO ProxyStructAlarmGroup
VAR_INPUT
	IOBJNUM : INT;
END_VAR
END_METHOD

METHOD GETPROXYHISTORICALALARMOBJECT : POINTER TO ProxyFbAlarmHistorical
VAR_INPUT
	XACTIVE : BOOL;
	IOBJNUM : INT;
END_VAR
END_METHOD

METHOD GETRECORDID : INT
END_METHOD

METHOD GETRECORDIDHISTORICAL : INT
END_METHOD

METHOD GETROWIDHISTORICALACTIVEALARMS
VAR_INPUT
	XFIRSTCALL : BOOL;
END_VAR
VAR_OUTPUT
	DWROWID : DWORD;
	LITS : LINT;
END_VAR
END_METHOD

METHOD GETROWTOREAD
VAR_OUTPUT
	DWROWIDLAST : DWORD;
	IROWCOUNT : INT;
END_VAR
END_METHOD

METHOD PRVCHECKALARMCLASS
VAR_INPUT
	PRECORDDATA : POINTER TO ProxyStructRecord;
END_VAR
END_METHOD

METHOD PRVCHECKALARMGROUP
VAR_INPUT
	PRECORDDATA : POINTER TO ProxyStructRecord;
END_VAR
END_METHOD

METHOD PRVGETALARMCLASSDESC : POINTER TO ProxyStructAlarmClass
VAR_INPUT
	PRECORDDATA : POINTER TO ProxyStructRecord;
	UICLASSID : UDINT;
END_VAR
END_METHOD

METHOD PRVGETALARMCLASSDESCBYNAME : POINTER TO ProxyStructAlarmClass
VAR_INPUT
	PRECORDDATA : POINTER TO ProxyStructRecord;
	SNAME : STRING;
END_VAR
END_METHOD

METHOD PRVGETALARMCONTAINER : POINTER TO AlarmContainer
VAR_INPUT
	DIOBJNUM : DINT;
	PSTRURECORD : POINTER TO ProxyStructRecord;
END_VAR
END_METHOD

METHOD PRVGETALARMDESC : POINTER TO ProxyStructAlarm
VAR_INPUT
	PRECORDDATA : POINTER TO ProxyStructRecord;
	UIALARMID : ALARM_ID;
	UDIGROUPID : UDINT;
END_VAR
END_METHOD

METHOD PRVGETALARMDESC2 : POINTER TO ProxyStructAlarm
VAR_INPUT
	PRECORDDATA : POINTER TO ProxyStructRecord;
	UDIALARMINTERNALID : UDINT;
	UDIGROUPID : UDINT;
END_VAR
END_METHOD

METHOD PRVGETALARMGROUPDESC : POINTER TO ProxyStructAlarmGroup
VAR_INPUT
	PSTRURECORD : POINTER TO ProxyStructRecord;
	UDIID : UDINT;
END_VAR
END_METHOD

METHOD PRVGETLOCK : RTS_IEC_HANDLE
VAR_INPUT
	ITASKID : INT;
END_VAR
END_METHOD

METHOD PRVGETPROXYACTIVEALARMOBJECT : IProxyAlarmObject
VAR_INPUT
	DIOBJNUM : DINT;
	PSTRURECORD : POINTER TO ProxyStructRecord;
END_VAR
END_METHOD

METHOD PRVGETRECORDDATA : POINTER TO ProxyStructRecord
VAR_INPUT
	IINDEX : INT;
END_VAR
END_METHOD

METHOD PRVPREPAREFORRESTART
END_METHOD

METHOD GETALARMCLASSESDESCRIPTION
VAR_INPUT
	PCLDESC : POINTER TO ARRAY [0..0] OF ProxyStructMonitorAlarmClassDesc;
	ISIZE : INT;
END_VAR
VAR_OUTPUT
	ICLCNT : INT;
END_VAR
END_METHOD

METHOD GETALARMGROUPSDESCRIPTION
VAR_INPUT
	PGRPDESC : POINTER TO ARRAY [0..0] OF ProxyStructMonitorAlarmGroupDesc;
	ISIZE : INT;
END_VAR
VAR_OUTPUT
	IGRPCNT : INT;
END_VAR
END_METHOD

METHOD GETALARMSDESCRIPTION
VAR_INPUT
	PALMDESC : POINTER TO ARRAY [0..0] OF ProxyStructMonitorAlarmDesc;
	DISIZE : DINT;
END_VAR
VAR_OUTPUT
	DIALMCNT : DINT;
END_VAR
END_METHOD

METHOD GETSTATISTICS : ProxyStructMonitor
VAR_INPUT
	IRECORD : INT;
END_VAR
END_METHOD

METHOD GETSTATISTICSSINGLEREQ : ProxyStructMonitorRequest
VAR_INPUT
	ITASKID : INT;
END_VAR
END_METHOD

METHOD PRVREADHISTALARMSPREELAB : SINT
VAR_INPUT
	IREQID : INT;
END_VAR
END_METHOD

METHOD PRVALARMOBJECTALLOC
VAR_INPUT
	PSTRURECORD : POINTER TO ProxyStructRecord;
END_VAR
END_METHOD

METHOD PRVALARMOBJECTFREE
VAR_INPUT
	PSTRURECORD : POINTER TO ProxyStructRecord;
END_VAR
END_METHOD

METHOD PRVALARMOBJECTSTUBSALLOC
VAR_INPUT
	PSTRURECORD : POINTER TO ProxyStructRecord;
END_VAR
END_METHOD

METHOD PRVALARMOBJECTSTUBSFREE
VAR_INPUT
	PSTRURECORD : POINTER TO ProxyStructRecord;
END_VAR
END_METHOD

METHOD PRVSTRUCTALARMCLASSDESCRIPTIONALLOC
VAR_INPUT
	PSTRURECORD : POINTER TO ProxyStructRecord;
END_VAR
END_METHOD

METHOD PRVSTRUCTALARMCLASSDESCRIPTIONFREE
VAR_INPUT
	PSTRURECORD : POINTER TO ProxyStructRecord;
END_VAR
END_METHOD

METHOD PRVSTRUCTALARMDESCRIPTIONALLOC
VAR_INPUT
	PSTRURECORD : POINTER TO ProxyStructRecord;
END_VAR
END_METHOD

METHOD PRVSTRUCTALARMDESCRIPTIONFREE
VAR_INPUT
	PSTRURECORD : POINTER TO ProxyStructRecord;
END_VAR
END_METHOD

METHOD PRVSTRUCTALARMGROUPDESCRIPTIONALLOC
VAR_INPUT
	PSTRURECORD : POINTER TO ProxyStructRecord;
END_VAR
END_METHOD

METHOD PRVSTRUCTALARMGROUPDESCRIPTIONFREE
VAR_INPUT
	PSTRURECORD : POINTER TO ProxyStructRecord;
END_VAR
END_METHOD

METHOD PRVGETENTRYTASKCALLTABLE : POINTER TO ProxyStructTaskCall
VAR_INPUT
	ITASKID : INT;
	ITABLE : INT;
END_VAR
END_METHOD

METHOD PRVPREPAREPRERUNTASKCALLTABLE
END_METHOD

METHOD PRVPREPARERUNTASKCALLTABLE
END_METHOD

(* ---- PROXYDATASOURCECHANNEL.fb ---- *)
FUNCTION_BLOCK PROXYDATASOURCECHANNEL
VAR
	M_ITFDATASOURCESMGR : IDatasources.IDatasourcesMgr;
	M_PSDSNAME : POINTER TO STRING;
	M_DIALARMNUM : DINT;
	M_IALARMCLASSNUM : INT;
	M_ILATCHVARSNUM : INT;
	M_ITFDATASOURCE : IDatasources.IDatasource2;
	M_IMAXALMGROUPS : INT;
	M_PSALMSTATETRANSCOUNTER : POINTER TO STRING;
	M_PALMSTATETRANSCOUNTER : __XWORD;
	M_TYPEALMSTATETRANSCOUNTER : TypeClass;
	M_XALMSTATETRANSCOUNTERISREG : BOOL;
	M_LIOLDSTATETRANSCOUNTERVALUE : LINT := -1;
	M_PSALMSTORAGECOUNTER : POINTER TO STRING;
	M_PALMSTORAGECOUNTER : __XWORD;
	M_TYPEALMSTORAGECOUNTER : TypeClass;
	M_XALMSTORAGECOUNTERISREG : BOOL;
	M_LIOLDSTORAGECOUNTERVALUE : LINT := -1;
	M_LIOLDSTORAGECOUNTERVALUE2 : LINT := -1;
	M_REQUESTBUILDERSETALMRECORD : RequestBuilderSetAlmRecord;
	M_REQUESTBUILDERRESALMRECORD : RequestBuilderResetAlmRecord;
	M_REQUESTBUILDERREADACTIVEALARMS : RequestBuilderReadActiveAlarms;
	M_REQUESTBUILDERGETALMCONFIG : RequestBuilderGetAlmConfig;
	M_REQUESTBUILDERGETALMCLASSCONFIG : RequestBuilderGetAlmClassConfig;
	M_REQUESTBUILDERACKALARMS : RequestBuilderAckAlarms;
	M_REQUESTBUILDERGETHISTORICALALMCONFIG : RequestBuilderGetHistoricalAlmConfig;
	M_REQUESTBUILDERREADHISTORICALALARMS : RequestBuilderReadHistoricalAlarms;
	M_REQUESTBUILDERREADHISTORICALACTIVEALARMS : RequestBuilderReadHistoricalActiveAlarms;
	M_REQUESTBUILDERCHANNELTEST : RequestBuilderChannelTest;
	M_REQUESTBUILDERCHANNELTEST2 : RequestBuilderChannelTest2;
	M_ITFPROXYCONSUMER : IProxyConsumer;
	M_ITFPROXYPROVIDER : IProxyProvider;
	M_ICURRREQUESTID : INT;
	M_ICOUNTTEST : INT;
	M_IERRORFROMDEV : INT;
	M_IHISTROWCOUNTREAD : INT;
	M_IHISTACTIVEROWCOUNTREAD : INT;
	M_IROWCOUNTREAD : INT;
	M_PFBREQUESTCALLED : POINTER TO RequestBuilderBase;
	M_XFIRSTCALL : BOOL := TRUE;
	M_LTLASTREADACTALM : LTIME;
	M_LTLASTREADHISTALM : LTIME;
	M_LTLASTREADHISTACTALM : LTIME;
	_SDEVICENAME : STRING;
	_ILATCHVARSNUM : INT;
	_IRECORDID : INT;
	_XHASSTORAGE : BOOL;
	_DWROWIDFIRST : DWORD;
	_DWROWIDLAST : DWORD;
	ALMSTATETRANSCOUNTERREGISTERED : BOOL;
	ALMSTORAGECOUNTERREGISTERED : BOOL;
	DEVICENAME : STRING;
	ERRORFROMDEVICE : INT;
	HASSTORAGE : BOOL;
	LATCHVARSNUM : INT;
	RECORDID : INT;
	ROWIDFIRST : DWORD;
	ROWIDLAST : DWORD;
	TESTVARIABLEVALUE : INT;
	TOTALARMNUM : DINT;
	TOTCLASSNUM : INT;
END_VAR
END_FUNCTION_BLOCK

METHOD SETPARAMS
VAR_INPUT
	PPARAM : POINTER TO ProxyStructDSChannelParam;
END_VAR
END_METHOD

METHOD GETCOUNTALARMSTOACKNOWLEDGE : INT
END_METHOD

METHOD GETNEXTALARMTOACKNOWLEDGE : BOOL
VAR_INPUT
	XFISRTENTRY : BOOL;
END_VAR
VAR_OUTPUT
	ALARMTOACKNOWLEDGE : AlarmToAcknowledge;
END_VAR
END_METHOD

METHOD GETPROXYALARMCLASSDESCRIPTIONOBJECT : POINTER TO ProxyStructAlarmClass
VAR_INPUT
	IOBJNUM : INT;
END_VAR
END_METHOD

METHOD GETPROXYALARMDESCRIPTIONOBJECT : POINTER TO ProxyStructAlarm
VAR_INPUT
	IOBJNUM : INT;
END_VAR
END_METHOD

METHOD GETPROXYALARMGROUPDESCRIPTIONOBJECT : POINTER TO ProxyStructAlarmGroup
VAR_INPUT
	IOBJNUM : INT;
END_VAR
END_METHOD

METHOD SETALARMMANAGERLIBVERSION
VAR_INPUT
	LIBVER : VERSION;
END_VAR
END_METHOD

METHOD SETALARMSCOUNT
VAR_INPUT
	DIVALUE : DINT;
END_VAR
END_METHOD

METHOD SETCLASSESCOUNT
VAR_INPUT
	IVALUE : INT;
END_VAR
END_METHOD

METHOD SETRECORDID
VAR_INPUT
	IVALUE : INT;
END_VAR
END_METHOD

METHOD GETALARMGROUP : STRING
VAR_INPUT
	IWHICHALARMGROUP : INT;
END_VAR
END_METHOD

METHOD GETALARMGROUPSNUM : INT
END_METHOD

METHOD SETVALUE
VAR_INPUT
	IVALUE : INT;
END_VAR
END_METHOD

METHOD GETVALUE : INT
END_METHOD

METHOD SETHASSTORAGE
VAR_INPUT
	XVALUE : BOOL;
END_VAR
END_METHOD

METHOD SETHISTACTIVEALARMSREAD
VAR_INPUT
	ICOUNT : INT;
END_VAR
END_METHOD

METHOD SETHISTALARMSREAD
VAR_INPUT
	DWROWIDLAST : DWORD;
	ICOUNT : INT;
	DISTORAGEROWSCOUNT : DINT;
	ISTORAGECLEAR : INT;
END_VAR
END_METHOD

METHOD SETROWIDS
VAR_INPUT
	DWROWIDFIRST : DWORD;
	DWROWIDLAST : DWORD;
END_VAR
END_METHOD

METHOD GETPROXYHISTORICALALARMOBJECT : POINTER TO ProxyFbAlarmHistorical
VAR_INPUT
	XACTIVE : BOOL;
	IOBJNUM : INT;
END_VAR
END_METHOD

METHOD GETRECORDIDHISTORICAL : INT
END_METHOD

METHOD GETROWIDHISTORICALACTIVEALARMS
VAR_INPUT
	XFIRSTCALL : BOOL;
END_VAR
VAR_OUTPUT
	DWROWID : DWORD;
	LITS : LINT;
END_VAR
END_METHOD

METHOD GETROWTOREAD
VAR_OUTPUT
	DWROWIDLAST : DWORD;
	IROWCOUNT : INT;
END_VAR
END_METHOD

METHOD ADDERROR
VAR_INPUT
	ITASKID : INT;
	UDIERROR : UDINT;
	SMSG : STRING;
END_VAR
END_METHOD

METHOD CLEANSTATISTICS : BOOL
VAR_INPUT
	ITASKID : INT;
END_VAR
END_METHOD

METHOD CYCLICCALL
END_METHOD

METHOD EXECUTEREQUEST : UDINT
VAR_INPUT
	ITASKID : INT;
	XLOCK : BOOL;
	HLOCK : RTS_IEC_HANDLE;
END_VAR
END_METHOD

METHOD GETALARMMESSAGETEXT : BOOL
VAR_INPUT
	ITFALARMMETAOBJECTSTUB5 : IAlarmMetaObjectStub5;
	IWHICHMESSAGE : INT;
	STRINGTYPE : __SYSTEM.TYPE_CLASS;
END_VAR
VAR_OUTPUT
	CBPMESSAGE : CharBufferPtr;
END_VAR
END_METHOD

METHOD GETALARMMESSAGETEXT2 : BOOL
VAR_INPUT
	STEXTLISTNAME : STRING;
	STEXTLISTINDEX : STRING;
	IWHICHMESSAGE : INT;
	STRINGTYPE : __SYSTEM.TYPE_CLASS;
END_VAR
VAR_OUTPUT
	CBPMESSAGE : CharBufferPtr;
END_VAR
END_METHOD

METHOD GETSTATISTICSSINGLEREQ : ProxyStructMonitorRequest
VAR_INPUT
	ITASKID : INT;
END_VAR
END_METHOD

METHOD INITIALIZE
VAR_INPUT
	ITFPROXYCONSUMER : IProxyConsumer;
	ITFPROXYPROVIDER : IProxyProvider;
	IMAXALMGROUPS : INT;
END_VAR
END_METHOD

METHOD ISCHANNELAVAILABLE : BOOL
END_METHOD

METHOD ISREQUESTEXECUTABLE : BOOL
VAR_INPUT
	ITASKID : INT;
	XTRYTOFORCE : BOOL;
END_VAR
END_METHOD

METHOD RESTART
END_METHOD

METHOD SETACTIVEALARMSCOUNT
VAR_INPUT
	DICOUNT : DINT;
END_VAR
END_METHOD

METHOD GETPROXYACTIVEALARMOBJECT : IProxyAlarmObject
VAR_INPUT
	DIOBJNUM : DINT;
END_VAR
END_METHOD

METHOD ERRORADDED
VAR_INPUT
	UDIERROR : UDINT;
	SMSG : STRING;
	STASKNAME : STRING;
END_VAR
END_METHOD

METHOD REQUESTCLOSED
VAR_INPUT
	IREQUESTID : INT;
END_VAR
END_METHOD

METHOD SETERRORFROMDEVICE
VAR_INPUT
	IERROR : INT;
END_VAR
END_METHOD

METHOD GETAPPLICATION : STRING
END_METHOD

METHOD GETDEVICENAME : STRING
END_METHOD

METHOD GETRECORDID : INT
END_METHOD

METHOD PRVGETALARMMESSAGETEXT
VAR_INPUT
	STEXTLISTNAME : STRING;
	STEXTLISTINDEX : STRING;
	IWHICHMESSAGE : INT;
	STRINGTYPE : __SYSTEM.TYPE_CLASS;
END_VAR
VAR_OUTPUT
	CBPMESSAGE : CharBufferPtr;
END_VAR
END_METHOD

METHOD PRVGETREQUESTBUILDERFB : POINTER TO RequestBuilderBase
VAR_INPUT
	ITASKID : INT;
END_VAR
END_METHOD

(* ---- PROXYFBALARMHISTORICAL.fb ---- *)
FUNCTION_BLOCK PROXYFBALARMHISTORICAL
VAR_INPUT
	M_DIHASTOREGISTERED : DINT;
	M_LATCHSTRINGS : ARRAY [1..MAX_LATCH_VARS] OF WSTRING;
	M_ROW : AlarmStorageRow;
END_VAR
VAR
	ALATCHVARIABLES : ARRAY [1..MAX_LATCH_VARS] OF LatchVariable;
	ALARMFB : Alarm;
END_VAR
END_FUNCTION_BLOCK

METHOD FB_INIT : BOOL
VAR_INPUT
	BINITRETAINS : BOOL;
	BINCOPYCODE : BOOL;
END_VAR
END_METHOD

(* ---- PROXYFBALARMMETAOBJECTSTUB.fb ---- *)
FUNCTION_BLOCK PROXYFBALARMMETAOBJECTSTUB
VAR_INPUT
	M_USILATCHVARSAVAIL : USINT;
END_VAR
VAR
	M_ALATCHVARIABLES : ARRAY [0..(MAX_LATCH_VARS - 1)] OF ValueTypeBundle;
	M_USICOUNTLATCHVARIABLES : USINT;
	M_UIID : ALARM_ID;
	M_UDIALARMGROUPINTERNALID : UDINT;
	M_LITIMESTAMPACKNOWLEDGE : AlarmManager_Interfaces.Timestamp;
	M_LITIMESTAMPACTIVE : AlarmManager_Interfaces.Timestamp;
	M_LITIMESTAMPINACTIVE : AlarmManager_Interfaces.Timestamp;
	M_LITIMESTAMPLAST : AlarmManager_Interfaces.Timestamp;
	M_IOFFSETACKNOWLEDGE : INT := -1;
	M_IOFFSETACTIVE : INT := -1;
	M_IOFFSETINACTIVE : INT := -1;
	M_IOFFSETLAST : INT := -1;
	M_ISTATE : INT;
	M_SALARMGROUP : STRING;
	M_STESTLISTNAME : STRING;
	M_SALARMCLASS : STRING;
	M_UDIALARMCLASSINTERNALID : UDINT;
	M_BYPRIORITY : BYTE;
	M_SALARMID : STRING;
	M_SPROXYNAME : STRING;
	M_CURRENTVALUE : ValueTypeBundle;
	M_TRIGGERVALUE : ValueTypeBundle;
	ALARMCLASSINTERNALID : UDINT;
	ALARMGROUPINTERNALID : UDINT;
	ALARMINTERNALID : UDINT;
	OFFSETACKNOWLEDGE : INT;
	OFFSETACTIVE : INT;
	OFFSETINACTIVE : INT;
	OFFSETLAST : INT;
	PROXYNAME : STRING;
END_VAR
END_FUNCTION_BLOCK

METHOD FB_EXIT : BOOL
VAR_INPUT
	BINCOPYCODE : BOOL;
END_VAR
END_METHOD

METHOD GETCHECKSUM : UDINT
END_METHOD

METHOD GETCURRENTVALUE : AlarmManagerInternal_Interfaces.ITypedValue
END_METHOD

METHOD SETACKNOWLEDGE
VAR_INPUT
	BACKNOWLEDGEMULTIPLE : BOOL;
END_VAR
END_METHOD

METHOD SWAPVALUES
END_METHOD

METHOD GETACKNOWLEDGE : BOOL
END_METHOD

METHOD GETACKNOWLEDGEMULTIPLE : BOOL
END_METHOD

METHOD GETALARMCLASS : STRING
END_METHOD

METHOD GETPRIORITY : BYTE
END_METHOD

METHOD GETSTRINGID : STRING
END_METHOD

METHOD GETTESTLISTNAME : STRING
END_METHOD

METHOD RESETACKNOWLEDGE
END_METHOD

METHOD SETALARMCLASS
VAR_INPUT
	SALARMCLASS : STRING;
END_VAR
END_METHOD

METHOD SETCURRENTVALUE
VAR_INPUT
	ITFTYPEDVALUECURRENT : AlarmManager_Interfaces.ITypedValue;
END_VAR
END_METHOD

METHOD SETPRIORITY
VAR_INPUT
	BYPRIORITY : BYTE;
END_VAR
END_METHOD

METHOD SETSTRINGID
VAR_INPUT
	SID : STRING;
END_VAR
END_METHOD

METHOD SETTESTLISTNAME
VAR_INPUT
	STESTLISTNAME : STRING;
END_VAR
END_METHOD

METHOD SETACKNOWLEDGE2
VAR_INPUT
	BACKNOWLEDGEMULTIPLE : BOOL;
END_VAR
END_METHOD

METHOD GETCOUNTLATCHVARIABLES : USINT
END_METHOD

METHOD GETLATCHVARVALUE : ITypedValue2
VAR_INPUT
	IWHICHLATCHVAR : INT;
END_VAR
END_METHOD

METHOD SETLATCHVARVALUE
VAR_INPUT
	IWHICHLATCHVAR : INT;
	ITFTYPEDVALUELATCHVAR : ITypedValue;
END_VAR
END_METHOD

METHOD SETCOUNTLATCHVARIABLES
VAR_INPUT
	USICOUNT : USINT;
END_VAR
END_METHOD

METHOD GETALARMGROUP : STRING
END_METHOD

METHOD GETID : AlarmManager_Interfaces.ALARM_ID
END_METHOD

METHOD GETLATCHVAR1VALUE : AlarmManager_Interfaces.ITypedValue
END_METHOD

METHOD GETLATCHVAR2VALUE : AlarmManager_Interfaces.ITypedValue
END_METHOD

METHOD GETSTATE : INT
END_METHOD

METHOD GETTIMESTAMPACKNOWLEDGE : AlarmManager_Interfaces.Timestamp
END_METHOD

METHOD GETTIMESTAMPACTIVE : AlarmManager_Interfaces.Timestamp
END_METHOD

METHOD GETTIMESTAMPINACTIVE : AlarmManager_Interfaces.Timestamp
END_METHOD

METHOD GETTIMESTAMPLAST : AlarmManager_Interfaces.Timestamp
END_METHOD

METHOD GETTRIGGERVALUE : AlarmManager_Interfaces.ITypedValue
END_METHOD

METHOD SETALARMGROUP
VAR_INPUT
	SALARMGROUP : STRING;
END_VAR
END_METHOD

METHOD SETID
VAR_INPUT
	UIID : AlarmManager_Interfaces.ALARM_ID;
END_VAR
END_METHOD

METHOD SETLATCHVAR1VALUE
VAR_INPUT
	ITFTYPEDVALUELATCHVAR1 : AlarmManager_Interfaces.ITypedValue;
END_VAR
END_METHOD

METHOD SETLATCHVAR2VALUE
VAR_INPUT
	ITFTYPEDVALUELATCHVAR2 : AlarmManager_Interfaces.ITypedValue;
END_VAR
END_METHOD

METHOD SETSTATE
VAR_INPUT
	ISTATE : INT;
END_VAR
END_METHOD

METHOD SETTIMESTAMPACKNOWLEDGE
VAR_INPUT
	LITIMESTAMPACKNOWLEDGE : AlarmManager_Interfaces.Timestamp;
END_VAR
END_METHOD

METHOD SETTIMESTAMPACTIVE
VAR_INPUT
	LITIMESTAMPACTIVE : AlarmManager_Interfaces.Timestamp;
END_VAR
END_METHOD

METHOD SETTIMESTAMPINACTIVE
VAR_INPUT
	LITIMESTAMPINACTIVE : AlarmManager_Interfaces.Timestamp;
END_VAR
END_METHOD

METHOD SETTIMESTAMPLAST
VAR_INPUT
	LITIMESTAMPLAST : AlarmManager_Interfaces.Timestamp;
END_VAR
END_METHOD

METHOD SETTRIGGERVALUE
VAR_INPUT
	ITFTYPEDVALUETRIGGER : AlarmManager_Interfaces.ITypedValue;
END_VAR
END_METHOD

(* ---- PROXYFBHISTACTIVEALARMSQUEUE.fb ---- *)
FUNCTION_BLOCK PROXYFBHISTACTIVEALARMSQUEUE
VAR
	M_PAALARM : POINTER TO ARRAY [0..10] OF POINTER TO ProxyStructHistoricalAlarmActive;
	M_DISZQUEUE : DINT;
	M_DISCANPOS : DINT;
	M_DICNTMAX : DINT;
	M_DICNT : DINT;
	M_DICNTAUX : DINT;
	SIZE_HIST_ACTIVE_ALARMS : INT := 50;
	EFFECTIVEREAD : DINT;
	QUEUESIZE : DINT;
END_VAR
END_FUNCTION_BLOCK

METHOD FB_EXIT : BOOL
VAR_INPUT
	BINCOPYCODE : BOOL;
END_VAR
END_METHOD

METHOD GETACTIVECOUNT : DINT
END_METHOD

METHOD GETAVAILABLEENTRIES : DINT
END_METHOD

METHOD GETLASTSTATE : AlarmState
VAR_INPUT
	DWROWID : DWORD;
END_VAR
END_METHOD

METHOD GETROWIDACTIVE
VAR_INPUT
	XFIRSTCALL : BOOL;
END_VAR
VAR_OUTPUT
	DWROWID : DWORD;
	LITS : LINT;
END_VAR
END_METHOD

METHOD GETROWIDLOCAL : DWORD
VAR_INPUT
	DWROWID : DWORD;
END_VAR
END_METHOD

METHOD INITIALIZE
END_METHOD

METHOD INSERT
VAR_INPUT
	SALM : ProxyStructHistoricalAlarmActive;
END_VAR
END_METHOD

METHOD ISPRESENTROWIDREMOTE : BOOL
VAR_INPUT
	DWROWID : DWORD;
END_VAR
END_METHOD

METHOD REMOVE
VAR_INPUT
	DWROWID : DWORD;
END_VAR
END_METHOD

METHOD SETLASTSTATE
VAR_INPUT
	DWROWID : DWORD;
	ESTATE : AlarmState;
END_VAR
END_METHOD

METHOD PRVHISTACTIVEENLARGE : BOOL
END_METHOD

(* ---- PROXYFBHISTALARMSROWQUEUE.fb ---- *)
FUNCTION_BLOCK PROXYFBHISTALARMSROWQUEUE
VAR
	M_PAHISTQUEUE : POINTER TO ARRAY [0..10] OF ProxyFbAlarmHistorical;
	M_ISZQUEUE : INT;
	MAXENTRIES : INT;
END_VAR
END_FUNCTION_BLOCK

METHOD FB_EXIT : BOOL
VAR_INPUT
	BINCOPYCODE : BOOL;
END_VAR
END_METHOD

METHOD GETAVAILABLEENTRIES : INT
END_METHOD

METHOD GETCOUNTTOREGISTER : INT
END_METHOD

METHOD GETITEM : POINTER TO ProxyFbAlarmHistorical
VAR_INPUT
	IOBJNUM : INT;
END_VAR
END_METHOD

METHOD INITIALIZE
VAR_INPUT
	SZQUEUE : INT;
END_VAR
END_METHOD

(* ---- REMOTEDEVICECOMPARER.fb ---- *)
FUNCTION_BLOCK REMOTEDEVICECOMPARER EXTENDS TSLastComparer
END_FUNCTION_BLOCK

METHOD COMPARE : INT
VAR_INPUT
	DIINDEXALARM1 : DINT;
	DIINDEXALARM2 : DINT;
END_VAR
END_METHOD

(* ---- REP_ACK_ALARMSTATEMACHINE.fb ---- *)
FUNCTION_BLOCK REP_ACK_ALARMSTATEMACHINE
END_FUNCTION_BLOCK

METHOD DOACKNOWLEDGE : AlarmState
VAR_INPUT
	ECURRENTSTATE : AlarmState;
END_VAR
VAR_OUTPUT
	ESTATETRANSITION : AlarmStateTransition;
END_VAR
END_METHOD

METHOD DOACTIVATE : AlarmState
VAR_INPUT
	ECURRENTSTATE : AlarmState;
END_VAR
END_METHOD

METHOD DODEACTIVATE : AlarmState
VAR_INPUT
	ECURRENTSTATE : AlarmState;
END_VAR
VAR_OUTPUT
	ESTATETRANSITION : AlarmStateTransition;
END_VAR
END_METHOD

(* ---- REP_ACK_ALARMSTATEMACHINE_NOCONFIRM.fb ---- *)
FUNCTION_BLOCK REP_ACK_ALARMSTATEMACHINE_NOCONFIRM EXTENDS Rep_Ack_AlarmStateMachine
END_FUNCTION_BLOCK

METHOD DOACKNOWLEDGE : AlarmState
VAR_INPUT
	ECURRENTSTATE : AlarmState;
END_VAR
VAR_OUTPUT
	ESTATETRANSITION : AlarmStateTransition;
END_VAR
END_METHOD

METHOD DODEACTIVATE : AlarmState
VAR_INPUT
	ECURRENTSTATE : AlarmState;
END_VAR
VAR_OUTPUT
	ESTATETRANSITION : AlarmStateTransition;
END_VAR
END_METHOD

(* ---- REP_ALARMSTATEMACHINE.fb ---- *)
FUNCTION_BLOCK REP_ALARMSTATEMACHINE
END_FUNCTION_BLOCK

METHOD DOACKNOWLEDGE : AlarmState
VAR_INPUT
	ECURRENTSTATE : AlarmState;
END_VAR
VAR_OUTPUT
	ESTATETRANSITION : AlarmStateTransition;
END_VAR
END_METHOD

METHOD DOACTIVATE : AlarmState
VAR_INPUT
	ECURRENTSTATE : AlarmState;
END_VAR
END_METHOD

METHOD DODEACTIVATE : AlarmState
VAR_INPUT
	ECURRENTSTATE : AlarmState;
END_VAR
VAR_OUTPUT
	ESTATETRANSITION : AlarmStateTransition;
END_VAR
END_METHOD

(* ---- REQUESTBUILDERACKALARMS.fb ---- *)
FUNCTION_BLOCK REQUESTBUILDERACKALARMS EXTENDS RequestBuilderBase
VAR
	M_ITFOWNSERVICEPROVIDER : IAckAlarmsServiceProvider;
	M_ITFOWNSERVICECONSUMER : IAckAlarmsServiceConsumer;
	COMPONENT : STRING := 'RequestBuilderReadActiveAlarms';
END_VAR
END_FUNCTION_BLOCK

METHOD BUILDANDENQUEUEV3REQUEST : UDINT
VAR_INPUT
	IREQUESTID : INT;
	ITFSERVICEPROVIDER : IServiceProvider;
	ITFSERVICECONSUMER : IServiceConsumer;
END_VAR
END_METHOD

METHOD FB_INIT : BOOL
VAR_INPUT
	BINITRETAINS : BOOL;
	BINCOPYCODE : BOOL;
END_VAR
END_METHOD

METHOD INITIALIZE
VAR_INPUT
	ITFDATASOURCE : IDatasources.IDatasource2;
	IMAXALMGROUPS : INT;
END_VAR
END_METHOD

METHOD BUILDREQUEST : UDINT
VAR_INPUT
	ITFSERVICEWRITER : CDSV3Prot.IServiceWriter;
	XHASTOSWAP : BOOL;
END_VAR
END_METHOD

METHOD GETSERVICE : UINT
END_METHOD

METHOD REQUESTFINISHED
VAR_INPUT
	REQUEST : IDatasources.ICustomRequest;
	RESPONSE : IDatasources.ICustomResponse;
	RESULT : SysTypes.RTS_IEC_RESULT;
END_VAR
END_METHOD

(* ---- REQUESTBUILDERBASE.fb ---- *)
FUNCTION_BLOCK REQUESTBUILDERBASE
VAR_INPUT
	M_REQUESTMONITOR : ProxyStructMonitorRequest;
	M_XLOCK : BOOL;
	M_HLOCK : RTS_IEC_HANDLE;
END_VAR
VAR
	M_ITFDATASOURCE : IDatasources.IDatasource2;
	M_ITFCDSV3REQUEST : IDatasources.ICDSV3Request;
	M_EBYTEORDER : IDatasources.ByteOrder := IDatasources.ByteOrder.Unknown;
	M_XHASTOSWAP : BOOL;
	M_ITFCDSV3REQUESTBUILDER : CDSV3Prot.ICDSV3RequestBuilder;
	M_ITFCUSTOMREQUESTCALLBACK : IDatasources.ICustomRequestCallback;
	M_PABYREQUESTBUFFER : POINTER TO BYTE;
	M_UDIREQUESTBUFFERSIZE : UDINT := MEM_SIZE_UNIT;
	M_ICURRREQUESTID : INT;
	M_IFBREQUESTID : INT;
	M_ITFSERVICECONSUMER : IServiceConsumer;
	M_LTSTARTTIME : LTIME;
	M_LTSTARTTIMEWAITANS : LTIME;
	M_UDIPREVERRCOUNT : UDINT;
	M_DURATION1 : Statistics_LTIME;
	M_IDURATIONSTATCNT : INT := 10;
	M_LTREQDURATIONLAST : LTIME;
	M_LTREQDURATIONAVG : LTIME;
	M_LTREQDURATIONMIN : LTIME;
	M_LTREQDURATIONMAX : LTIME;
	M_LTREQDURATIONBUILDREQ : LTIME;
	M_LTREQDURATIONWAITANS : LTIME;
	M_LTREQDURATIONELABANS : LTIME;
	M_SCOMPONENT : STRING := 'RequestBuilderBase';
	M_LOCKRESULT : RTS_IEC_RESULT := Errors.ERR_FAILED;
	MEM_SIZE_UNIT : UDINT := 256;
	MEM_SIZE_UNIT_GRP : UDINT := (MEM_SIZE_UNIT * 4);
	ISERRORPRESENT : BOOL;
END_VAR
END_FUNCTION_BLOCK

METHOD ADDERROR
VAR_INPUT
	UDIERROR : UDINT;
	SMSG : STRING;
END_VAR
END_METHOD

METHOD BUILDANDENQUEUEV3REQUEST : UDINT
VAR_INPUT
	IREQUESTID : INT;
	ITFSERVICEPROVIDER : IServiceProvider;
	ITFSERVICECONSUMER : IServiceConsumer;
END_VAR
END_METHOD

METHOD FB_EXIT : BOOL
VAR_INPUT
	BINCOPYCODE : BOOL;
END_VAR
END_METHOD

METHOD GETSTATISTICSDATA
END_METHOD

METHOD INITIALIZE
VAR_INPUT
	ITFDATASOURCE : IDatasources.IDatasource2;
	IMAXALMGROUPS : INT;
END_VAR
END_METHOD

METHOD BUILDREQUEST : UDINT
VAR_INPUT
	ITFSERVICEWRITER : CDSV3Prot.IServiceWriter;
	XHASTOSWAP : BOOL;
END_VAR
END_METHOD

METHOD GETDATABUFFER : POINTER TO BYTE
END_METHOD

METHOD GETDATABUFFERSIZE : UDINT
END_METHOD

METHOD GETSERVICE : UINT
END_METHOD

METHOD GETSERVICEGROUP : UINT
END_METHOD

METHOD REQUESTENQUEUED : UDINT
END_METHOD

METHOD SETTARGETBYTEORDER
VAR_INPUT
	EBYTEORDER : IDatasources.ByteOrder;
END_VAR
END_METHOD

METHOD REQUESTFINISHED
VAR_INPUT
	REQUEST : IDatasources.ICustomRequest;
	RESPONSE : IDatasources.ICustomResponse;
	RESULT : SysTypes.RTS_IEC_RESULT;
END_VAR
END_METHOD

METHOD PROTAFTERBUILDREQUEST
END_METHOD

METHOD PROTAFTERREQUEST
VAR_INPUT
	ITFSERVICECONSUMER : IServiceConsumer;
END_VAR
END_METHOD

METHOD PROTBEFOREANSELAB
END_METHOD

METHOD PROTBEFOREREQUEST
VAR_INPUT
	IREQUESTID : INT;
END_VAR
END_METHOD

METHOD PROTBUILDANDENQUEUEV3REQUEST : UDINT
END_METHOD

METHOD PROTRELEASEREQUEST
END_METHOD

(* ---- REQUESTBUILDERCHANNELTEST.fb ---- *)
FUNCTION_BLOCK REQUESTBUILDERCHANNELTEST EXTENDS RequestBuilderBase
VAR
	M_ITFOWNSERVICEPROVIDER : IChannelTestServiceProvider;
	M_ITFOWNSERVICECONSUMER : IChannelTestServiceConsumer;
	COMPONENT : STRING := 'RequestBuilderChannelTest';
END_VAR
END_FUNCTION_BLOCK

METHOD BUILDANDENQUEUEV3REQUEST : UDINT
VAR_INPUT
	IREQUESTID : INT;
	ITFSERVICEPROVIDER : IServiceProvider;
	ITFSERVICECONSUMER : IServiceConsumer;
END_VAR
END_METHOD

METHOD FB_INIT : BOOL
VAR_INPUT
	BINITRETAINS : BOOL;
	BINCOPYCODE : BOOL;
END_VAR
END_METHOD

METHOD INITIALIZE
VAR_INPUT
	ITFDATASOURCE : IDatasources.IDatasource2;
	IMAXALMGROUPS : INT;
END_VAR
END_METHOD

METHOD BUILDREQUEST : UDINT
VAR_INPUT
	ITFSERVICEWRITER : CDSV3Prot.IServiceWriter;
	XHASTOSWAP : BOOL;
END_VAR
END_METHOD

METHOD GETSERVICE : UINT
END_METHOD

METHOD REQUESTFINISHED
VAR_INPUT
	REQUEST : IDatasources.ICustomRequest;
	RESPONSE : IDatasources.ICustomResponse;
	RESULT : SysTypes.RTS_IEC_RESULT;
END_VAR
END_METHOD

(* ---- REQUESTBUILDERCHANNELTEST2.fb ---- *)
FUNCTION_BLOCK REQUESTBUILDERCHANNELTEST2 EXTENDS RequestBuilderChannelTest
VAR
	COMPONENT2 : STRING := 'RequestBuilderChannelTest2';
END_VAR
END_FUNCTION_BLOCK

METHOD FB_INIT : BOOL
VAR_INPUT
	BINITRETAINS : BOOL;
	BINCOPYCODE : BOOL;
END_VAR
END_METHOD

METHOD INITIALIZE
VAR_INPUT
	ITFDATASOURCE : IDatasources.IDatasource2;
	IMAXALMGROUPS : INT;
END_VAR
END_METHOD

(* ---- REQUESTBUILDERGETALMCLASSCONFIG.fb ---- *)
FUNCTION_BLOCK REQUESTBUILDERGETALMCLASSCONFIG EXTENDS RequestBuilderBase
VAR
	M_ITFOWNSERVICEPROVIDER : IAlmConfigServiceProvider;
	M_ITFOWNSERVICECONSUMER : IAlmConfigServiceConsumer;
	COMPONENT : STRING := 'RequestBuilderGetAlmClassConfig';
END_VAR
END_FUNCTION_BLOCK

METHOD BUILDANDENQUEUEV3REQUEST : UDINT
VAR_INPUT
	IREQUESTID : INT;
	ITFSERVICEPROVIDER : IServiceProvider;
	ITFSERVICECONSUMER : IServiceConsumer;
END_VAR
END_METHOD

METHOD FB_INIT : BOOL
VAR_INPUT
	BINITRETAINS : BOOL;
	BINCOPYCODE : BOOL;
END_VAR
END_METHOD

METHOD INITIALIZE
VAR_INPUT
	ITFDATASOURCE : IDatasources.IDatasource2;
	IMAXALMGROUPS : INT;
END_VAR
END_METHOD

METHOD BUILDREQUEST : UDINT
VAR_INPUT
	ITFSERVICEWRITER : CDSV3Prot.IServiceWriter;
	XHASTOSWAP : BOOL;
END_VAR
END_METHOD

METHOD GETSERVICE : UINT
END_METHOD

METHOD REQUESTFINISHED
VAR_INPUT
	REQUEST : IDatasources.ICustomRequest;
	RESPONSE : IDatasources.ICustomResponse;
	RESULT : SysTypes.RTS_IEC_RESULT;
END_VAR
END_METHOD

(* ---- REQUESTBUILDERGETALMCONFIG.fb ---- *)
FUNCTION_BLOCK REQUESTBUILDERGETALMCONFIG EXTENDS RequestBuilderBase
VAR
	M_ITFOWNSERVICEPROVIDER : IAlmConfigServiceProvider;
	M_ITFOWNSERVICECONSUMER : IAlmConfigServiceConsumer;
	COMPONENT : STRING := 'RequestBuilderGetAlmConfig';
END_VAR
END_FUNCTION_BLOCK

METHOD BUILDANDENQUEUEV3REQUEST : UDINT
VAR_INPUT
	IREQUESTID : INT;
	ITFSERVICEPROVIDER : IServiceProvider;
	ITFSERVICECONSUMER : IServiceConsumer;
END_VAR
END_METHOD

METHOD FB_INIT : BOOL
VAR_INPUT
	BINITRETAINS : BOOL;
	BINCOPYCODE : BOOL;
END_VAR
END_METHOD

METHOD INITIALIZE
VAR_INPUT
	ITFDATASOURCE : IDatasources.IDatasource2;
	IMAXALMGROUPS : INT;
END_VAR
END_METHOD

METHOD BUILDREQUEST : UDINT
VAR_INPUT
	ITFSERVICEWRITER : CDSV3Prot.IServiceWriter;
	XHASTOSWAP : BOOL;
END_VAR
END_METHOD

METHOD GETSERVICE : UINT
END_METHOD

METHOD REQUESTFINISHED
VAR_INPUT
	REQUEST : IDatasources.ICustomRequest;
	RESPONSE : IDatasources.ICustomResponse;
	RESULT : SysTypes.RTS_IEC_RESULT;
END_VAR
END_METHOD

(* ---- REQUESTBUILDERGETHISTORICALALMCONFIG.fb ---- *)
FUNCTION_BLOCK REQUESTBUILDERGETHISTORICALALMCONFIG EXTENDS RequestBuilderBase
VAR
	M_ITFOWNSERVICEPROVIDER : IHistoricAlmServiceProvider;
	M_ITFOWNSERVICECONSUMER : IHistoricAlmServiceConsumer;
	COMPONENT : STRING := 'RequestBuilderGetHistoricalAlmConfig';
END_VAR
END_FUNCTION_BLOCK

METHOD BUILDANDENQUEUEV3REQUEST : UDINT
VAR_INPUT
	IREQUESTID : INT;
	ITFSERVICEPROVIDER : IServiceProvider;
	ITFSERVICECONSUMER : IServiceConsumer;
END_VAR
END_METHOD

METHOD FB_INIT : BOOL
VAR_INPUT
	BINITRETAINS : BOOL;
	BINCOPYCODE : BOOL;
END_VAR
END_METHOD

METHOD INITIALIZE
VAR_INPUT
	ITFDATASOURCE : IDatasources.IDatasource2;
	IMAXALMGROUPS : INT;
END_VAR
END_METHOD

METHOD BUILDREQUEST : UDINT
VAR_INPUT
	ITFSERVICEWRITER : CDSV3Prot.IServiceWriter;
	XHASTOSWAP : BOOL;
END_VAR
END_METHOD

METHOD GETSERVICE : UINT
END_METHOD

METHOD REQUESTFINISHED
VAR_INPUT
	REQUEST : IDatasources.ICustomRequest;
	RESPONSE : IDatasources.ICustomResponse;
	RESULT : SysTypes.RTS_IEC_RESULT;
END_VAR
END_METHOD

(* ---- REQUESTBUILDERREADACTIVEALARMS.fb ---- *)
FUNCTION_BLOCK REQUESTBUILDERREADACTIVEALARMS EXTENDS RequestBuilderBase
VAR
	M_ITFOWNSERVICEPROVIDER : IReadActiveAlarmsServiceProvider;
	M_ITFOWNSERVICECONSUMER : IReadActiveAlarmsServiceConsumer;
	COMPONENT : STRING := 'RequestBuilderReadActiveAlarms';
END_VAR
END_FUNCTION_BLOCK

METHOD BUILDANDENQUEUEV3REQUEST : UDINT
VAR_INPUT
	IREQUESTID : INT;
	ITFSERVICEPROVIDER : IServiceProvider;
	ITFSERVICECONSUMER : IServiceConsumer;
END_VAR
END_METHOD

METHOD FB_INIT : BOOL
VAR_INPUT
	BINITRETAINS : BOOL;
	BINCOPYCODE : BOOL;
END_VAR
END_METHOD

METHOD INITIALIZE
VAR_INPUT
	ITFDATASOURCE : IDatasources.IDatasource2;
	IMAXALMGROUPS : INT;
END_VAR
END_METHOD

METHOD BUILDREQUEST : UDINT
VAR_INPUT
	ITFSERVICEWRITER : CDSV3Prot.IServiceWriter;
	XHASTOSWAP : BOOL;
END_VAR
END_METHOD

METHOD GETSERVICE : UINT
END_METHOD

METHOD REQUESTFINISHED
VAR_INPUT
	REQUEST : IDatasources.ICustomRequest;
	RESPONSE : IDatasources.ICustomResponse;
	RESULT : SysTypes.RTS_IEC_RESULT;
END_VAR
END_METHOD

(* ---- REQUESTBUILDERREADHISTORICALACTIVEALARMS.fb ---- *)
FUNCTION_BLOCK REQUESTBUILDERREADHISTORICALACTIVEALARMS EXTENDS RequestBuilderBase
VAR
	M_ITFOWNSERVICEPROVIDER : IHistoricAlmServiceProvider;
	M_ITFOWNSERVICECONSUMER : IHistoricAlmServiceConsumer;
	COMPONENT : STRING := 'RequestBuilderReadHistoricalActiveAlarms';
END_VAR
END_FUNCTION_BLOCK

METHOD BUILDANDENQUEUEV3REQUEST : UDINT
VAR_INPUT
	IREQUESTID : INT;
	ITFSERVICEPROVIDER : IServiceProvider;
	ITFSERVICECONSUMER : IServiceConsumer;
END_VAR
END_METHOD

METHOD FB_INIT : BOOL
VAR_INPUT
	BINITRETAINS : BOOL;
	BINCOPYCODE : BOOL;
END_VAR
END_METHOD

METHOD INITIALIZE
VAR_INPUT
	ITFDATASOURCE : IDatasources.IDatasource2;
	IMAXALMGROUPS : INT;
END_VAR
END_METHOD

METHOD BUILDREQUEST : UDINT
VAR_INPUT
	ITFSERVICEWRITER : CDSV3Prot.IServiceWriter;
	XHASTOSWAP : BOOL;
END_VAR
END_METHOD

METHOD GETSERVICE : UINT
END_METHOD

METHOD REQUESTFINISHED
VAR_INPUT
	REQUEST : IDatasources.ICustomRequest;
	RESPONSE : IDatasources.ICustomResponse;
	RESULT : SysTypes.RTS_IEC_RESULT;
END_VAR
END_METHOD

(* ---- REQUESTBUILDERREADHISTORICALALARMS.fb ---- *)
FUNCTION_BLOCK REQUESTBUILDERREADHISTORICALALARMS EXTENDS RequestBuilderBase
VAR
	M_ITFOWNSERVICEPROVIDER : IHistoricAlmServiceProvider;
	M_ITFOWNSERVICECONSUMER : IHistoricAlmServiceConsumer;
	COMPONENT : STRING := 'RequestBuilderReadHistoricalAlarms';
END_VAR
END_FUNCTION_BLOCK

METHOD BUILDANDENQUEUEV3REQUEST : UDINT
VAR_INPUT
	IREQUESTID : INT;
	ITFSERVICEPROVIDER : IServiceProvider;
	ITFSERVICECONSUMER : IServiceConsumer;
END_VAR
END_METHOD

METHOD FB_INIT : BOOL
VAR_INPUT
	BINITRETAINS : BOOL;
	BINCOPYCODE : BOOL;
END_VAR
END_METHOD

METHOD INITIALIZE
VAR_INPUT
	ITFDATASOURCE : IDatasources.IDatasource2;
	IMAXALMGROUPS : INT;
END_VAR
END_METHOD

METHOD BUILDREQUEST : UDINT
VAR_INPUT
	ITFSERVICEWRITER : CDSV3Prot.IServiceWriter;
	XHASTOSWAP : BOOL;
END_VAR
END_METHOD

METHOD GETSERVICE : UINT
END_METHOD

METHOD REQUESTFINISHED
VAR_INPUT
	REQUEST : IDatasources.ICustomRequest;
	RESPONSE : IDatasources.ICustomResponse;
	RESULT : SysTypes.RTS_IEC_RESULT;
END_VAR
END_METHOD

(* ---- REQUESTBUILDERRESETALMRECORD.fb ---- *)
FUNCTION_BLOCK REQUESTBUILDERRESETALMRECORD EXTENDS RequestBuilderBase
VAR
	M_ITFOWNSERVICEPROVIDER : IAlmRecordServiceProvider;
	M_ITFOWNSERVICECONSUMER : IAlmRecordServiceConsumer;
	COMPONENT : STRING := 'RequestBuilderResetAlmRecord';
END_VAR
END_FUNCTION_BLOCK

METHOD BUILDANDENQUEUEV3REQUEST : UDINT
VAR_INPUT
	IREQUESTID : INT;
	ITFSERVICEPROVIDER : IServiceProvider;
	ITFSERVICECONSUMER : IServiceConsumer;
END_VAR
END_METHOD

METHOD FB_INIT : BOOL
VAR_INPUT
	BINITRETAINS : BOOL;
	BINCOPYCODE : BOOL;
END_VAR
END_METHOD

METHOD INITIALIZE
VAR_INPUT
	ITFDATASOURCE : IDatasources.IDatasource2;
	IMAXALMGROUPS : INT;
END_VAR
END_METHOD

METHOD BUILDREQUEST : UDINT
VAR_INPUT
	ITFSERVICEWRITER : CDSV3Prot.IServiceWriter;
	XHASTOSWAP : BOOL;
END_VAR
END_METHOD

METHOD GETSERVICE : UINT
END_METHOD

METHOD REQUESTFINISHED
VAR_INPUT
	REQUEST : IDatasources.ICustomRequest;
	RESPONSE : IDatasources.ICustomResponse;
	RESULT : SysTypes.RTS_IEC_RESULT;
END_VAR
END_METHOD

(* ---- REQUESTBUILDERSETALMRECORD.fb ---- *)
FUNCTION_BLOCK REQUESTBUILDERSETALMRECORD EXTENDS RequestBuilderBase
VAR
	M_ITFOWNSERVICEPROVIDER : IAlmRecordServiceProvider;
	M_ITFOWNSERVICECONSUMER : IAlmRecordServiceConsumer;
	COMPONENT : STRING := 'RequestBuilderSetAlmRecord';
END_VAR
END_FUNCTION_BLOCK

METHOD BUILDANDENQUEUEV3REQUEST : UDINT
VAR_INPUT
	IREQUESTID : INT;
	ITFSERVICEPROVIDER : IServiceProvider;
	ITFSERVICECONSUMER : IServiceConsumer;
END_VAR
END_METHOD

METHOD FB_INIT : BOOL
VAR_INPUT
	BINITRETAINS : BOOL;
	BINCOPYCODE : BOOL;
END_VAR
END_METHOD

METHOD INITIALIZE
VAR_INPUT
	ITFDATASOURCE : IDatasources.IDatasource2;
	IMAXALMGROUPS : INT;
END_VAR
END_METHOD

METHOD BUILDREQUEST : UDINT
VAR_INPUT
	ITFSERVICEWRITER : CDSV3Prot.IServiceWriter;
	XHASTOSWAP : BOOL;
END_VAR
END_METHOD

METHOD GETSERVICE : UINT
END_METHOD

METHOD REQUESTFINISHED
VAR_INPUT
	REQUEST : IDatasources.ICustomRequest;
	RESPONSE : IDatasources.ICustomResponse;
	RESULT : SysTypes.RTS_IEC_RESULT;
END_VAR
END_METHOD

(* ---- ROWIDCOMPARER.fb ---- *)
FUNCTION_BLOCK ROWIDCOMPARER EXTENDS AbstractComparer
END_FUNCTION_BLOCK

METHOD COMPARE : INT
VAR_INPUT
	DIINDEXALARM1 : DINT;
	DIINDEXALARM2 : DINT;
END_VAR
END_METHOD

(* ---- RUNTIMEEVENTLISTENER.fb ---- *)
FUNCTION_BLOCK RUNTIMEEVENTLISTENER
VAR
	_HPREPAREDOWNLOADEVENT : RTS_IEC_HANDLE := Events.Invalid_Handle;
	_HPREPAREDOWNLOADEVENTINTERFACE : RTS_IEC_HANDLE := Events.Invalid_Handle;
	_HPREPARESTOPEVENT : RTS_IEC_HANDLE := Events.Invalid_Handle;
	_HPREPARESTOPEVENTINTERFACE : RTS_IEC_HANDLE := Events.Invalid_Handle;
END_VAR
END_FUNCTION_BLOCK

METHOD EVENTCALLBACK : UDINT
VAR_INPUT
	PEVENTPARAM : POINTER TO EventParam;
END_VAR
END_METHOD

METHOD FB_EXIT : BOOL
VAR_INPUT
	BINCOPYCODE : BOOL;
END_VAR
END_METHOD

METHOD FB_INIT : BOOL
VAR_INPUT
	BINITRETAINS : BOOL;
	BINCOPYCODE : BOOL;
END_VAR
END_METHOD

METHOD PRVISOURAPPLICATIONBEFOREDELETE : BOOL
VAR_INPUT
	PAPPDELETEEVENTPARAM : POINTER TO CmPApp.EVTPARAM_CmpAppStop;
END_VAR
END_METHOD

METHOD PRVISOURAPPLICATIONBEFOREDOWNLOAD : BOOL
VAR_INPUT
	PAPPEVENTPARAM : POINTER TO CmPApp.EVTPARAM_CmpApp;
END_VAR
END_METHOD

(* ---- SERIALIZERDATABLOCK.fb ---- *)
FUNCTION_BLOCK SERIALIZERDATABLOCK
VAR_INPUT
	M_PBYBUFFER : POINTER TO BYTE;
	M_UDIBUFFERSIZE : UDINT;
END_VAR
VAR
	M_SERIALIZINGALARMMETAOBJECTSTUB : SerializingAlarmMetaObjectStub;
	M_ICOUNTROWS : INT;
	ERROR : UINT;
END_VAR
END_FUNCTION_BLOCK

METHOD GETALARMMETAOBJECTSTUB : IAlarmMetaObjectStub3
VAR_INPUT
	IROW : INT;
	IOFFSET : INT;
END_VAR
END_METHOD

METHOD GETCOUNTROWS : INT
END_METHOD

METHOD SETCOUNTROWS : BOOL
VAR_INPUT
	ICOUNT : INT;
END_VAR
END_METHOD

METHOD HASALARMS : BOOL
END_METHOD

METHOD SETTOTALCOUNTROWS : BOOL
VAR_INPUT
	DICOUNT : DINT;
END_VAR
END_METHOD

(* ---- SERIALIZINGALARMMETAOBJECTSTUB.fb ---- *)
FUNCTION_BLOCK SERIALIZINGALARMMETAOBJECTSTUB
VAR_INPUT
	M_PBYBUFFER : POINTER TO BYTE;
	M_UDIBUFFERSIZE : UDINT;
	M_UDIOFFSET : UDINT;
	M_XOVERFLOW : BOOL;
END_VAR
VAR
	S_OFFSET_TIMESTAMP_LAST : UDINT := 0;
	S_OFFSET_TIMESTAMP_ACTIVE : UDINT := (8 + s_OFFSET_TIMESTAMP_LAST);
	S_OFFSET_TIMESTAMP_INACTIVE : UDINT := (8 + s_OFFSET_TIMESTAMP_ACTIVE);
	S_OFFSET_TIMESTAMP_ACKNOWLEDGE : UDINT := (8 + s_OFFSET_TIMESTAMP_INACTIVE);
	S_OFFSET_TRIGGER_VALUE : UDINT := (8 + s_OFFSET_TIMESTAMP_ACKNOWLEDGE);
	S_OFFSET_LATCH1_VALUE : UDINT := (8 + s_OFFSET_TRIGGER_VALUE);
	S_OFFSET_LATCH2_VALUE : UDINT := (8 + s_OFFSET_LATCH1_VALUE);
	S_OFFSET_ALARMGROUP_ID : UDINT := (8 + s_OFFSET_LATCH2_VALUE);
	S_OFFSET_ALARM_ID : UDINT := (4 + s_OFFSET_ALARMGROUP_ID);
	S_OFFSET_STATE : UDINT := (4 + s_OFFSET_ALARM_ID);
	S_OFFSET_TRIGGER_VALUE_TYPE : UDINT := (1 + s_OFFSET_STATE);
	S_OFFSET_LATCH1_TYPE : UDINT := (1 + s_OFFSET_TRIGGER_VALUE_TYPE);
	S_OFFSET_LATCH2_TYPE : UDINT := (1 + s_OFFSET_LATCH1_TYPE);
	SIZE_LATCH2_TYPE : UDINT := 1;
	SIZE : UDINT;
END_VAR
END_FUNCTION_BLOCK

METHOD INITIALIZE
END_METHOD

METHOD SETALARM
VAR_INPUT
	PALARM : POINTER TO Alarm;
END_VAR
END_METHOD

METHOD SETLATCHVAR1VALUE
VAR_INPUT
	ITFTYPEDVALUELATCHVAR1 : ITypedValue;
END_VAR
END_METHOD

METHOD SETLATCHVAR2VALUE
VAR_INPUT
	ITFTYPEDVALUELATCHVAR2 : ITypedValue;
END_VAR
END_METHOD

METHOD SETSTATE
VAR_INPUT
	ISTATE : INT;
END_VAR
END_METHOD

METHOD SETTIMESTAMPACKNOWLEDGE
VAR_INPUT
	LITIMESTAMPACKNOWLEDGE : Timestamp;
END_VAR
END_METHOD

METHOD SETTIMESTAMPACTIVE
VAR_INPUT
	LITIMESTAMPACTIVE : Timestamp;
END_VAR
END_METHOD

METHOD SETTIMESTAMPINACTIVE
VAR_INPUT
	LITIMESTAMPINACTIVE : Timestamp;
END_VAR
END_METHOD

METHOD SETTIMESTAMPLAST
VAR_INPUT
	LITIMESTAMPLAST : Timestamp;
END_VAR
END_METHOD

METHOD SETTRIGGERVALUE
VAR_INPUT
	ITFTYPEDVALUETRIGGER : ITypedValue;
END_VAR
END_METHOD

METHOD GETALARM : POINTER TO Alarm
END_METHOD

METHOD GETALARMGROUP : STRING
END_METHOD

METHOD GETCHECKSUM : UDINT
END_METHOD

METHOD GETCURRENTVALUE : ITypedValue
END_METHOD

METHOD GETID : ALARM_ID
END_METHOD

METHOD GETLATCHVAR1VALUE : ITypedValue
END_METHOD

METHOD GETLATCHVAR2VALUE : ITypedValue
END_METHOD

METHOD GETSTATE : INT
END_METHOD

METHOD GETTIMESTAMPACKNOWLEDGE : Timestamp
END_METHOD

METHOD GETTIMESTAMPACTIVE : Timestamp
END_METHOD

METHOD GETTIMESTAMPINACTIVE : Timestamp
END_METHOD

METHOD GETTIMESTAMPLAST : Timestamp
END_METHOD

METHOD GETTRIGGERVALUE : ITypedValue
END_METHOD

METHOD SETACKNOWLEDGE
VAR_INPUT
	BACKNOWLEDGEMULTIPLE : BOOL;
END_VAR
END_METHOD

METHOD SETALARMGROUP
VAR_INPUT
	SALARMGROUP : STRING;
END_VAR
END_METHOD

METHOD SETCURRENTLREALVALUE
VAR_INPUT
	LRVALUE : LREAL;
END_VAR
END_METHOD

METHOD SETCURRENTVALUE
VAR_INPUT
	ITFTYPEDVALUECURRENT : ITypedValue;
END_VAR
END_METHOD

METHOD SETID
VAR_INPUT
	UIID : ALARM_ID;
END_VAR
END_METHOD

(* ---- SQLITEDATABASEACCESS.fb ---- *)
FUNCTION_BLOCK SQLITEDATABASEACCESS EXTENDS AbstractDatabaseAccess
VAR
	M_CONTEXT : SQLiteDatabaseAccessContext;
	M_ITFALARMSTORAGEMANAGER : IAlarmStorageManager;
	M_ISUPPORTEDVERSION : INT := -1;
	M_XBYTEORDERGET : BOOL;
END_VAR
END_FUNCTION_BLOCK

METHOD SETALARMSTORAGEMANAGER
VAR_INPUT
	ITFALARMSTORAGEMANAGER : IAlarmStorageManager;
END_VAR
END_METHOD

METHOD GETNUMBEROFLATCHVARIABLES : USINT
END_METHOD

METHOD GETROOTPAGE : CAA.IDENT
VAR_INPUT
	EWHICHALARMSTORAGEOBJECT : EAlarmStorageObject;
END_VAR
END_METHOD

METHOD ISONLYONEALARMCLASSSELECTED : BOOL
END_METHOD

METHOD ISONLYONEALARMGROUPSELECTED : BOOL
END_METHOD

METHOD PREPAREDATABASEACCESS : STO.ERROR
END_METHOD

METHOD TBLALARMCURSORCLOSE : STO.ERROR
VAR_INPUT
	EERRORFROMPREVIOUSPROCESSING : STO.ERROR;
END_VAR
END_METHOD

METHOD TBLALARMCURSORMOVE : STO.ERROR
VAR_INPUT
	EDIRECTION : STO.DIRECTION;
END_VAR
VAR_OUTPUT
	XEOF : BOOL;
END_VAR
END_METHOD

METHOD TBLALARMCURSOROPEN : STO.ERROR
VAR_INPUT
	FILTERCRITERIA : REFERENCE TO VisuFbAlarmFilterCriteria;
END_VAR
END_METHOD

METHOD TBLALARMCURSOROPEN2 : STO.ERROR
VAR_INPUT
	IDINDEX : CAA.IDENT;
END_VAR
END_METHOD

METHOD TBLALARMCURSORSETPOSITION : STO.ERROR
VAR_INPUT
	FILTERCRITERIA : REFERENCE TO VisuFbAlarmFilterCriteria;
	BROWIDVALID : BOOL;
	DIROWID : DINT;
END_VAR
END_METHOD

METHOD TBLALARMGETLATCHVARTYPE : STO.ERROR
VAR_INPUT
	IDWHICHCOLUMN : CAA.IDENT;
	USIWHICHLATCHVAR : USINT;
END_VAR
VAR_OUTPUT
	BYTYPE : BYTE;
	XNULL : BOOL;
END_VAR
END_METHOD

METHOD TBLALARMGETLATCHVARVALUE : STO.ERROR
VAR_INPUT
	IDWHICHCOLUMN : CAA.IDENT;
	USIWHICHLATCHVAR : USINT;
END_VAR
VAR_OUTPUT
	LIVALUE : LINT;
	XNULL : BOOL;
END_VAR
END_METHOD

METHOD TBLALARMGETMINMAXROWIDS : BOOL
VAR_OUTPUT
	IDROWMIN : LINT;
	IDROWMAX : LINT;
	EERROR : STO.ERROR;
END_VAR
END_METHOD

METHOD TBLALARMGETROWCOUNT : CAA.COUNT
VAR_OUTPUT
	EERROR : STO.ERROR;
END_VAR
END_METHOD

METHOD TBLALARMGETTIMESTAMPVALUE : LINT
VAR_INPUT
	IDWHICHCOLUMN : CAA.IDENT;
END_VAR
VAR_OUTPUT
	EERROR : STO.ERROR;
END_VAR
END_METHOD

METHOD TBLALARMGET_DINT : STO.ERROR
VAR_INPUT
	IDWHICHCOLUMN : CAA.IDENT;
	IWHICHCOLUMN : INT;
END_VAR
VAR_OUTPUT
	DIVALUE : DINT;
	XNULL : BOOL;
END_VAR
END_METHOD

METHOD TBLALARMGET_LINT : STO.ERROR
VAR_INPUT
	IDWHICHCOLUMN : CAA.IDENT;
	IWHICHCOLUMN : INT;
END_VAR
VAR_OUTPUT
	LIVALUE : LINT;
	XNULL : BOOL;
END_VAR
END_METHOD

METHOD TBLALARMGET_SINT : STO.ERROR
VAR_INPUT
	IDWHICHCOLUMN : CAA.IDENT;
	IWHICHCOLUMN : INT;
END_VAR
VAR_OUTPUT
	SIVALUE : SINT;
	XNULL : BOOL;
END_VAR
END_METHOD

METHOD TBLALARMISNOTEMPTY : BOOL
VAR_OUTPUT
	EERROR : STO.ERROR;
END_VAR
END_METHOD

METHOD TBLALARMROWGETCURRENT : STO.ERROR
END_METHOD

METHOD TBLALARMROWGETCURRENTID : DINT
END_METHOD

METHOD TBLALARMROWISVALID : BOOL
END_METHOD

METHOD TBLALARMROWRELEASE : STO.ERROR
VAR_INPUT
	EERRORFROMPREVIOUSPROCESSING : STO.ERROR;
END_VAR
END_METHOD

METHOD TBLALARMROWSELECT : STO.ERROR
VAR_INPUT
	IDROW : CAA.IDENT;
	XDOERRORHANDLING : BOOL;
END_VAR
END_METHOD

METHOD TBLALARMTABLECLOSE : STO.ERROR
END_METHOD

METHOD TBLALARMTABLEISOPEN : BOOL
END_METHOD

METHOD TBLALARMTABLEOPEN : STO.ERROR
VAR_INPUT
	XREADONLY : BOOL;
END_VAR
END_METHOD

METHOD TBLLATCHVARSTRINGSCLOSEIFNEEDED : STO.ERROR
VAR_INPUT
	EERRORFROMPREVIOUSPROCESSING : STO.ERROR;
END_VAR
END_METHOD

METHOD TBLLATCHVARSTRINGSCURSORSEARCHROWID : STO.ERROR
VAR_INPUT
	LIROWID : LINT;
END_VAR
END_METHOD

METHOD TBLLATCHVARSTRINGSGET_TEXT : STO.ERROR
VAR_INPUT
	IDWHICHCOLUMN : CAA.IDENT;
	IWHICHCOLUMN : INT;
END_VAR
VAR_OUTPUT
	XNULL : BOOL;
END_VAR
VAR_IN_OUT
	TXTVALUE : STO.TEXT;
END_VAR
END_METHOD

METHOD TBLLATCHVARSTRINGSOPENIFNEEDED : STO.ERROR
END_METHOD

METHOD TBLLATCHVARSTRINGSROWGETCURRENT : STO.ERROR
END_METHOD

METHOD TBLLATCHVARSTRINGSROWRELEASE : STO.ERROR
VAR_INPUT
	EERRORFROMPREVIOUSPROCESSING : STO.ERROR;
END_VAR
END_METHOD

METHOD TEXTCOPYTOSTRING : STO.ERROR
VAR_INPUT
	XFREE : BOOL;
END_VAR
VAR_IN_OUT
	TXTVALUE : STO.TEXT;
	SVALUE : STRING(1);
	SZVALUE : CAA.SIZE;
END_VAR
END_METHOD

METHOD TEXTCOPYTOWSTRING : STO.ERROR
VAR_INPUT
	XFREE : BOOL;
END_VAR
VAR_IN_OUT
	TXTVALUE : STO.TEXT;
	WSVALUE : WSTRING(1);
	SZVALUE : CAA.SIZE;
END_VAR
END_METHOD

METHOD TRANSACTIONBEGIN : STO.ERROR
VAR_INPUT
	XREADONLY : BOOL;
END_VAR
END_METHOD

METHOD TRANSACTIONBEGINFAILED : BOOL
END_METHOD

METHOD TRANSACTIONEND
VAR_INPUT
	EERRORFROMPREVIOUSPROCESSING : STO.ERROR;
END_VAR
END_METHOD

METHOD TBLALARMGET_INT : STO.ERROR
VAR_INPUT
	IDWHICHCOLUMN : CAA.IDENT;
	IWHICHCOLUMN : INT;
END_VAR
VAR_OUTPUT
	IVALUE : INT;
	XNULL : BOOL;
END_VAR
END_METHOD

METHOD TBLVERSIONGETCURRENT : STO.ERROR
VAR_OUTPUT
	IVERSION : INT;
END_VAR
END_METHOD

METHOD GETRELEVANTFILTERDATA
VAR_OUTPUT
	EDBBYTEORDER : EAlarmByteOrder;
END_VAR
END_METHOD

METHOD TBLALARMCURSORSEARCHROWID : STO.ERROR
VAR_INPUT
	IDROW : DINT;
END_VAR
END_METHOD

METHOD TBLGETBYTEORDER : STO.ERROR
VAR_OUTPUT
	EBYTEORDER : EAlarmByteOrder;
END_VAR
END_METHOD

METHOD TBLVERSIONGETCURRENT2 : STO.ERROR
VAR_OUTPUT
	IVERSION : INT;
	EDBUSED : EDBType;
END_VAR
END_METHOD

METHOD TBLALARMGETCOMMENTVALUE : STO.ERROR
VAR_INPUT
	IDWHICHCOLUMN : CAA.IDENT;
	IWHICHCOLUMN : INT;
END_VAR
VAR_OUTPUT
	XNULL : BOOL;
END_VAR
VAR_IN_OUT
	WSVALUE : WSTRING(2000);
END_VAR
END_METHOD

(* ---- STANDARDALARMCONFIGURATION.fb ---- *)
FUNCTION_BLOCK STANDARDALARMCONFIGURATION
VAR
	M_PAITFALARMGROUPS : POINTER TO ARRAY [0..0] OF IAlarmGroup;
	M_ICOUNTALARMGROUPS : INT;
	M_PAITFALARMCLASSES : POINTER TO ARRAY [0..0] OF IAlarmClass;
	M_ICOUNTALARMCLASSES : INT;
	M_XVARIABLESREGISTERED : BOOL;
	M_XFIRST : BOOL;
	M_XPLACEHOLDANALYZED : BOOL;
	M_LTSTARTTIME : LTIME;
	M_DATABASESIZELIMIT : DatabaseSizeLimit;
	M_XDATABASESIZELIMITBLOCKED : BOOL;
	_XRAISEDMOREALARMSTHANSTORAGELIMITREPORTED : BOOL;
	_XCLEARHISTORY : BOOL;
	_XKEEPACTIVEALARMS : BOOL;
	M_DICTALARMTEMPLATEINSTANCES : AlarmInstanceDictionary;
	M_SZAPPNAME : STRING(CmpApp.GlobalConstants.MAX_LEN_APPLNAME);
	DATABASESIZELIMIT : IDatabaseSizeLimit;
	TOTALROWSTOINSERT : UDINT;
END_VAR
END_FUNCTION_BLOCK

METHOD FB_EXIT : BOOL
VAR_INPUT
	BINCOPYCODE : BOOL;
END_VAR
END_METHOD

METHOD FB_INIT : BOOL
VAR_INPUT
	BINITRETAINS : BOOL;
	BINCOPYCODE : BOOL;
END_VAR
END_METHOD

METHOD FINDALARMBYID : IAlarm
VAR_INPUT
	USIALARMGROUPID : ALARMGROUP_ID;
	UIALARMID : ALARM_ID;
END_VAR
END_METHOD

METHOD REGISTERVARIABLES
END_METHOD

METHOD ADDTOINSTANCEDICTIONARY : BOOL
VAR_INPUT
	PINSTANCE : POINTER TO BYTE;
	PSTALARMTEMPLATENAME : POINTER TO STRING;
	UDIALARMGROUPID : UDINT;
	UITEMPLATEALARMSOFFSET : UINT;
	UITEMPLATEALARMSLENGTH : UINT;
	UITEMPLATEEVENTSOFFSET : UINT;
	UITEMPLATEEVENTSLENGTH : UINT;
END_VAR
END_METHOD

METHOD CLEARINSTANCEDICTIONARY : BOOL
END_METHOD

METHOD GETALARMFROMDICTIONARY : IAlarm8
VAR_INPUT
	PINSTANCE : POINTER TO BYTE;
	UDIALARMID : REFERENCE TO ALARM_ID;
	STALARMTEMPLATENAME : REFERENCE TO STRING;
END_VAR
VAR_OUTPUT
	USIALARMGROUPID : ALARMGROUP_ID;
	UIALARMID : ALARM_ID;
END_VAR
END_METHOD

METHOD CREATEALARMSTORAGETASK
VAR_INPUT
	STSTORAGETASKGROUPNAME : REFERENCE TO STRING;
END_VAR
END_METHOD

METHOD INITSTORAGETASKINFO
VAR_INPUT
	ITASKPRIORITY : INT;
	DWINTERVAL : DWORD;
END_VAR
END_METHOD

METHOD ACKNOWLEDGEALL
END_METHOD

METHOD ACKNOWLEDGEALLOFGROUP
VAR_INPUT
	USIALARMGROUPID : ALARMGROUP_ID;
END_VAR
END_METHOD

METHOD ACKNOWLEDGEONEOFGROUP
VAR_INPUT
	USIALARMGROUPID : ALARMGROUP_ID;
	UIALARMID : ALARM_ID;
END_VAR
END_METHOD

METHOD CYCLICCALL
END_METHOD

METHOD FINDALARM : POINTER TO Alarm
VAR_INPUT
	SALARMGROUP : STRING;
	UIALARMID : ALARM_ID;
END_VAR
END_METHOD

METHOD FINDALARMCLASS : IAlarmClass
VAR_INPUT
	UDIID : UDINT;
END_VAR
END_METHOD

METHOD FINDALARMGROUP : IAlarmGroup
VAR_INPUT
	UDIID : UDINT;
END_VAR
END_METHOD

METHOD GETSTORAGE : IDatabaseFileAlarmStorage
END_METHOD

METHOD HASSTORAGE : BOOL
END_METHOD

METHOD RAISEEVENT : BOOL
VAR_INPUT
	EVENT : AlarmEvent;
END_VAR
END_METHOD

METHOD DETERMINERELEVANTALARMS : UDINT
VAR_INPUT
	ITFALARMFILTERCRITERIA : IAlarmFilterCriteria;
	PARRITFRELEVANTALARMS : POINTER TO ARRAY [0..0] OF IAlarm;
	IOFFSET : INT;
END_VAR
END_METHOD

METHOD FINDALARMGROUPBYNAME : IAlarmGroup
VAR_INPUT
	SALARMGROUP : STRING;
END_VAR
END_METHOD

METHOD FINDALARMCLASSBYNAME : IAlarmClass
VAR_INPUT
	SALARMCLASS : STRING;
END_VAR
END_METHOD

METHOD RAISEEVENT2 : BOOL
VAR_INPUT
	EVENT : AlarmEvent;
END_VAR
VAR_OUTPUT
	ITFALARM : IAlarm;
END_VAR
END_METHOD

METHOD GETALARMGROUPS : POINTER TO ARRAY [0..0] OF IAlarmGroup
VAR_OUTPUT
	IALARMGROUPCOUNT : INT;
END_VAR
END_METHOD

METHOD FINDALARMCLASSCOUNT : INT
END_METHOD

METHOD CLEARHISTORY : BOOL
VAR_INPUT
	XKEEPACTIVEALARMS : BOOL;
END_VAR
END_METHOD

METHOD ACKNOWLEDGEALLOFGROUPWITHCOMMENT
VAR_INPUT
	USIALARMGROUPID : ALARMGROUP_ID;
END_VAR
VAR_IN_OUT
	WSCOMMENT : WSTRING;
	WSUSERID : WSTRING;
END_VAR
END_METHOD

METHOD ACKNOWLEDGEALLWITHCOMMENT
VAR_IN_OUT
	WSCOMMENT : WSTRING;
	WSUSERID : WSTRING;
END_VAR
END_METHOD

METHOD ACKNOWLEDGEONEOFGROUPWITHCOMMENT
VAR_INPUT
	USIALARMGROUPID : ALARMGROUP_ID;
	UIALARMID : ALARM_ID;
END_VAR
VAR_IN_OUT
	WSCOMMENT : WSTRING;
	WSUSERID : WSTRING;
END_VAR
END_METHOD

METHOD SETCOMMENT : UDINT
VAR_INPUT
	USIALARMGROUPID : ALARMGROUP_ID;
	UIALARMID : ALARM_ID;
END_VAR
VAR_IN_OUT
	WSCOMMENT : WSTRING;
	WSUSERID : WSTRING;
END_VAR
END_METHOD

METHOD TRAVERSEALLALARMSOFALLALARMGROUPS
VAR_INPUT
	ITFALARMTRAVERSALCONSUMER : IAlarmTraversalConsumer;
END_VAR
END_METHOD

METHOD TRAVERSEALLCLASSES
VAR_INPUT
	ITFALARMTRAVERSALCONSUMER : IAlarmTraversalConsumer;
END_VAR
END_METHOD

METHOD NOTIFYREINITDONE
END_METHOD

METHOD CLEARALLALARMHISTORYENTRIESIFWISHED : BOOL
VAR_INPUT
	ITFDATABASEFILEALARMSTORAGE : IDatabaseFileAlarmStorage;
END_VAR
END_METHOD

METHOD CLEARONLYHISTORYOFINACTIVEALARMS : BOOL
END_METHOD

METHOD PRVACKNOWLEDGE
VAR_INPUT
	PAALARMS : POINTER TO ARRAY [0..0] OF Alarm;
	IALARMCOUNT : INT;
	UIALARMID : ALARM_ID;
	XACKALL : BOOL;
	PWSCOMMENT : POINTER TO WSTRING;
	PWSUSER : POINTER TO WSTRING;
END_VAR
END_METHOD

METHOD PRVCHECKSETACKNOWLEDGE
VAR_INPUT
	INDEX : INT;
	UIALARMID : ALARM_ID;
	XACKALL : BOOL;
	PWSCOMMENT : POINTER TO WSTRING;
	PWSUSER : POINTER TO WSTRING;
END_VAR
END_METHOD

METHOD PRVCREATEALARMSTORAGEMETADATAFILE
END_METHOD

METHOD PRVDETERMINERELEVANTALARMS : UDINT
VAR_INPUT
	PAALARMS : POINTER TO ARRAY [0..0] OF Alarm;
	IALARMCOUNT : INT;
	ITFALARMFILTERCRITERIA : IAlarmFilterCriteria;
	PARRITFRELEVANTALARMS : POINTER TO ARRAY [0..0] OF IAlarm;
	IOFFSET : INT;
END_VAR
END_METHOD

METHOD PRVINITIALIZEALARMCONFIGURATION
END_METHOD

METHOD PRVTRYGETCURRENTROW : BOOL
VAR_OUTPUT
	CURRENTROW : AlarmStorageRow;
END_VAR
END_METHOD

METHOD PRVTSTPLACEHOLDERS : BOOL
VAR_INPUT
	ALARM : REFERENCE TO Alarm;
END_VAR
END_METHOD

METHOD PRVWITHBRACKETS : STRING
VAR_INPUT
	SSTRING : STRING;
END_VAR
END_METHOD

METHOD PRVWITHOPENINGBRACKET : STRING
VAR_INPUT
	SSTRING : STRING;
END_VAR
END_METHOD

(* ---- STANDARDALARMCONFIGURATIONREMOTE.fb ---- *)
FUNCTION_BLOCK STANDARDALARMCONFIGURATIONREMOTE
VAR_INPUT
	M_PAITFPROXY : POINTER TO ARRAY [0..10] OF IProxy;
	M_IPROXYNUM : INT;
END_VAR
VAR
	M_SIALREADYSCAN : SINT := -1;
	PROXYNUM : INT;
END_VAR
END_FUNCTION_BLOCK

METHOD CYCLICCALL
END_METHOD

METHOD GETACTIVEALARMS
VAR_INPUT
	PASNAME : POINTER TO ARRAY [0..10] OF STRING;
	IGROUPCOUNT : INT;
	FILTERCRITERIA : REFERENCE TO VisuFbAlarmFilterCriteria;
	ITFALARMDATABLOCK : IAlarmDataBlockBaseDINT;
END_VAR
VAR_IN_OUT
	DISTUBPROG : DINT;
END_VAR
END_METHOD

METHOD GETALARMCLASSDESC : BOOL
VAR_INPUT
	SPROXYNAME : STRING;
	UDIID : UDINT;
END_VAR
VAR_OUTPUT
	SDESC : ProxyStructAlarmClassDesc;
END_VAR
END_METHOD

METHOD GETALARMCLASSDESCBYNAME : BOOL
VAR_INPUT
	SPROXYNAME : STRING;
	SCLASSNAME : STRING;
END_VAR
VAR_OUTPUT
	SDESC : ProxyStructAlarmClassDesc;
END_VAR
END_METHOD

METHOD GETALARMDESC : BOOL
VAR_INPUT
	SPROXYNAME : STRING;
	UDIALMID : UDINT;
	UDIGRPID : UDINT;
END_VAR
VAR_OUTPUT
	SDESC : ProxyStructAlarmDesc;
END_VAR
END_METHOD

METHOD GETALARMDISPLAYOPTIONS : BOOL
VAR_INPUT
	ITFALARMMETAOBJECTSTUB5 : IAlarmMetaObjectStub5;
	REFDISPLAYOPTIONS : REFERENCE TO DisplayOptions;
END_VAR
VAR_OUTPUT
	XVALID : BOOL;
	SCLASSREMAP : STRING;
END_VAR
END_METHOD

METHOD GETALARMGROUPDESC : BOOL
VAR_INPUT
	SPROXYNAME : STRING;
	UDIID : UDINT;
END_VAR
VAR_OUTPUT
	SDESC : ProxyStructAlarmGroupDesc;
END_VAR
END_METHOD

METHOD GETALARMGROUPDESCBYNAME : BOOL
VAR_INPUT
	SPROXYNAME : STRING;
	SGRPNAME : STRING;
END_VAR
VAR_OUTPUT
	SDESC : ProxyStructAlarmGroupDesc;
END_VAR
END_METHOD

METHOD GETALARMMESSAGE : BOOL
VAR_INPUT
	ITFALARMMETAOBJECTSTUB5 : IAlarmMetaObjectStub5;
	IWHICHMESSAGE : INT;
	REFCHARBUFFERSTRING : REFERENCE TO CharBufferString;
	STRINGTYPE : __SYSTEM.TYPE_CLASS;
END_VAR
END_METHOD

METHOD GETALARMMESSAGE2 : BOOL
VAR_INPUT
	SNAME : STRING;
	STEXTLISTNAME : STRING;
	STEXTLISTINDEX : STRING;
	IWHICHMESSAGE : INT;
	STRINGTYPE : __SYSTEM.TYPE_CLASS;
END_VAR
VAR_OUTPUT
	MESSAGE : CharBufferPtr;
END_VAR
END_METHOD

METHOD GETPROXY : IProxy
VAR_INPUT
	SNAME : STRING;
END_VAR
END_METHOD

METHOD GETSTORAGE : IDatabaseFileAlarmStorage
END_METHOD

METHOD HASSTORAGE : BOOL
END_METHOD

METHOD REGISTERUSERCLIENT : BOOL
VAR_INPUT
	IINDEX : INT;
END_VAR
VAR_OUTPUT
	ITFPROXY : IProxy;
END_VAR
END_METHOD

METHOD SETALARMSTOACK
VAR_INPUT
	ITFALARMDATABLOCK : IAlarmDataBlockBase2;
END_VAR
END_METHOD

METHOD REMOTEDEVICEREACHED
VAR_INPUT
	ROW : REFERENCE TO AlarmStorageRow;
	XFIRST : BOOL;
	IVERSION : INT;
END_VAR
END_METHOD

METHOD PRVGETPROXY : IProxy
VAR_INPUT
	SNAME : STRING;
END_VAR
END_METHOD

METHOD GETPROXYALARMCLASSESDESCRIPTION : BOOL
VAR_INPUT
	SNAME : STRING;
	PCLDESC : POINTER TO ARRAY [0..0] OF ProxyStructMonitorAlarmClassDesc;
	ISIZE : INT;
END_VAR
VAR_OUTPUT
	ICLCNT : INT;
END_VAR
END_METHOD

METHOD GETPROXYALARMGROUPSDESCRIPTION : BOOL
VAR_INPUT
	SNAME : STRING;
	PGRPDESC : POINTER TO ARRAY [0..0] OF ProxyStructMonitorAlarmGroupDesc;
	ISIZE : INT;
END_VAR
VAR_OUTPUT
	IGRPCNT : INT;
END_VAR
END_METHOD

METHOD GETPROXYALARMSDESCRIPTION : BOOL
VAR_INPUT
	SNAME : STRING;
	PALMDESC : POINTER TO ARRAY [0..0] OF ProxyStructMonitorAlarmDesc;
	DISIZE : DINT;
END_VAR
VAR_OUTPUT
	DIALMCNT : DINT;
END_VAR
END_METHOD

METHOD GETPROXYSTATISTICS : BOOL
VAR_INPUT
	SNAME : STRING;
END_VAR
VAR_OUTPUT
	STRUCTMONITOR : ProxyStructMonitor;
END_VAR
END_METHOD

METHOD GETPROXYSTATISTICSSINGLEACTIVITY : BOOL
VAR_INPUT
	SNAME : STRING;
	ITASKID : INT;
END_VAR
VAR_OUTPUT
	STRUCTMONITOR : ProxyStructMonitorRequest;
END_VAR
END_METHOD

(* ---- STANDARDALARMHANDLER.fb ---- *)
FUNCTION_BLOCK STANDARDALARMHANDLER
VAR
	M_AITFALARMCONFIGURATIONS : ARRAY [0..(MAX_COUNT_CONFIG - 1)] OF IAlarmConfiguration;
	M_ICOUNTCONFIGURATIONS : INT := 0;
	M_AITFALARMCONFIGURATIONSREM : ARRAY [0..(MAX_COUNT_CONFIG - 1)] OF IAlarmConfigurationRemote;
	M_ICOUNTCONFIGURATIONSREM : INT := 0;
	M_ALARMMANAGERCLIENTINFOSTRUCTVECTOR : AlarmManagerClientInfoStructVector;
	M_DIALARMSTATETRANSITIONCOUNTERPREVIOUSCALL : DINT;
	M_DIALARMSTORAGECOUNTERPREVIOUSCALL : DINT;
	M_ITFSTORAGETODELETE : IDatabaseFileAlarmStorage;
	M_XSTART : BOOL := TRUE;
	M_XFIRSTCYCLEAFTERDOWNLOAD : BOOL := TRUE;
	MAX_COUNT_CONFIG : BYTE := 2;
	ALARMCONFIGURATIONCOUNT : INT;
	ISREADY : BOOL;
END_VAR
END_FUNCTION_BLOCK

METHOD FB_EXIT : BOOL
VAR_INPUT
	BINCOPYCODE : BOOL;
END_VAR
END_METHOD

METHOD FB_INIT : BOOL
VAR_INPUT
	BINITRETAINS : BOOL;
	BINCOPYCODE : BOOL;
END_VAR
END_METHOD

METHOD FINDALARM : POINTER TO Alarm
VAR_INPUT
	SALARMGROUP : STRING;
	UIALARMID : ALARM_ID;
END_VAR
END_METHOD

METHOD FINDALARMCLASSBYNAME : IAlarmClass
VAR_INPUT
	SALARMCLASS : STRING;
END_VAR
END_METHOD

METHOD FINDALARMCLASSCOUNTALL : INT
END_METHOD

METHOD FINDALARMGROUPBYNAME : IAlarmGroup
VAR_INPUT
	SALARMGROUP : STRING;
END_VAR
END_METHOD

METHOD FINDALARMGROUPBYNAMEALL : IAlarmGroup
VAR_INPUT
	SALARMGROUP : STRING;
END_VAR
END_METHOD

METHOD REREGISTERCLIENTS
END_METHOD

METHOD TRAVERSEALLALARMSOFALLALARMCONFIGURATIONS
VAR_INPUT
	ITFALARMTRAVERSALCONSUMER : IAlarmTraversalConsumer;
END_VAR
END_METHOD

METHOD TRAVERSEALLCLASSESOFALLALARMCONFIGURATIONS
VAR_INPUT
	ITFALARMTRAVERSALCONSUMER : IAlarmTraversalConsumer;
END_VAR
END_METHOD

METHOD ALLOCBYTES : POINTER TO BYTE
VAR_INPUT
	UXISIZE : __UXINT;
END_VAR
END_METHOD

METHOD ALLOCFBALARMCLASSADAPTER : POINTER TO AlarmClassAdapter
END_METHOD

METHOD ALLOCFBALARMGROUPADAPTER : POINTER TO AlarmGroupAdapter
END_METHOD

METHOD ALLOCVALUETYPEBUNDLE : POINTER TO ValueTypeBundle
END_METHOD

METHOD ACKNOWLEDGEALL
END_METHOD

METHOD ACKNOWLEDGEALLOFGROUP
VAR_INPUT
	USIALARMGROUPID : ALARMGROUP_ID;
END_VAR
END_METHOD

METHOD ACKNOWLEDGEONEOFGROUP
VAR_INPUT
	USIALARMGROUPID : ALARMGROUP_ID;
	UIALARMID : ALARM_ID;
END_VAR
END_METHOD

METHOD CYCLICCALL
END_METHOD

METHOD FINDALARMCLASS : IAlarmClass
VAR_INPUT
	UDIID : UDINT;
END_VAR
END_METHOD

METHOD FINDALARMGROUP : IAlarmGroup
VAR_INPUT
	UDIID : UDINT;
END_VAR
END_METHOD

METHOD GETSTORAGE : IDatabaseFileAlarmStorage
END_METHOD

METHOD HASSTORAGE : BOOL
END_METHOD

METHOD RAISEEVENT : BOOL
VAR_INPUT
	USIALARMGROUPID : ALARMGROUP_ID;
	UIALARMID : ALARM_ID;
END_VAR
END_METHOD

METHOD REGISTERALARMCONFIGURATION
VAR_INPUT
	ITFALARMCONFIGURATION : IAlarmConfiguration;
END_VAR
END_METHOD

METHOD GETACTIVEALARMS : UDINT
VAR_INPUT
	ITFALARMMANAGERCLIENT : IAlarmManagerClient;
END_VAR
VAR_OUTPUT
	PARRITFACTIVEALARMS : POINTER TO ARRAY [0..0] OF IAlarm;
	ICOUNTACTIVEALARMS : INT;
END_VAR
END_METHOD

METHOD GETALARMSFROMSTORAGE : UDINT
VAR_INPUT
	ITFALARMMANAGERCLIENT : IAlarmManagerClient;
	ISKIPROWS : INT;
END_VAR
VAR_OUTPUT
	ICOUNTROWS : INT;
END_VAR
VAR_IN_OUT
	BROWIDVALID : BOOL;
	DIROWID : DINT;
END_VAR
END_METHOD

METHOD GETCOUNTALARMSFROMSTORAGE : DINT
VAR_INPUT
	ITFALARMMANAGERCLIENT : IAlarmManagerClient;
END_VAR
VAR_OUTPUT
	UDIRESULT : UDINT;
END_VAR
END_METHOD

METHOD REGISTERCLIENT : UDINT
VAR_INPUT
	ITFALARMMANAGERCLIENT : IAlarmManagerClient;
	PARRITFALARMSFROMHISTORY : POINTER TO ARRAY [0..0] OF IAlarm2;
	ICOUNTALARMSFROMHISTORY : INT;
END_VAR
END_METHOD

METHOD UNREGISTERCLIENT : UDINT
VAR_INPUT
	ITFALARMMANAGERCLIENT : IAlarmManagerClient;
END_VAR
END_METHOD

METHOD UNREGISTERALARMCONFIGURATION
VAR_INPUT
	ITFALARMCONFIGURATION : IAlarmConfiguration;
END_VAR
END_METHOD

METHOD REGISTERALARMSTATECHANGEDLISTENER : BOOL
VAR_INPUT
	ITFALARMSTATECHANGEDLISTENER : IAlarmStateChangedListener;
END_VAR
END_METHOD

METHOD GETALARMCONFIGURATION : IAlarmConfiguration
VAR_INPUT
	IPOS : INT;
END_VAR
END_METHOD

METHOD ACKNOWLEDGEALLOFGROUPWITHCOMMENT
VAR_INPUT
	USIALARMGROUPID : ALARMGROUP_ID;
END_VAR
VAR_IN_OUT
	WSCOMMENT : WSTRING;
	WSUSERID : WSTRING;
END_VAR
END_METHOD

METHOD ACKNOWLEDGEALLWITHCOMMENT
VAR_IN_OUT
	WSCOMMENT : WSTRING;
	WSUSERID : WSTRING;
END_VAR
END_METHOD

METHOD ACKNOWLEDGEONEOFGROUPWITHCOMMENT
VAR_INPUT
	USIALARMGROUPID : ALARMGROUP_ID;
	UIALARMID : ALARM_ID;
END_VAR
VAR_IN_OUT
	WSCOMMENT : WSTRING;
	WSUSERID : WSTRING;
END_VAR
END_METHOD

METHOD SETCOMMENT : UDINT
VAR_INPUT
	USIALARMGROUPID : ALARMGROUP_ID;
	UIALARMID : ALARM_ID;
END_VAR
VAR_IN_OUT
	WSCOMMENT : WSTRING;
	WSUSERID : WSTRING;
END_VAR
END_METHOD

METHOD GETINSTANCEALARM : IAlarm8
VAR_INPUT
	PFBINSTANCE : POINTER TO BYTE;
	UITEMPLATEALARMID : ALARM_ID;
END_VAR
VAR_OUTPUT
	USIALARMGROUPID : ALARMGROUP_ID;
	UIALARMID : ALARM_ID;
END_VAR
END_METHOD

METHOD GETINSTANCEALARMBYNAME : IAlarm8
VAR_INPUT
	PFBINSTANCE : POINTER TO BYTE;
	UITEMPLATEALARMID : ALARM_ID;
	STALARMTEMPLATENAME : STRING(255);
END_VAR
VAR_OUTPUT
	USIALARMGROUPID : ALARMGROUP_ID;
	UIALARMID : ALARM_ID;
END_VAR
END_METHOD

METHOD RAISEEVENTALARMINSTANCE : BOOL
VAR_INPUT
	PFBINSTANCE : POINTER TO BYTE;
	UITEMPLATEALARMID : ALARM_ID;
END_VAR
END_METHOD

METHOD RAISEEVENTALARMINSTANCEBYNAME : BOOL
VAR_INPUT
	PFBINSTANCE : POINTER TO BYTE;
	UITEMPLATEALARMID : ALARM_ID;
	STALARMTEMPLATENAME : STRING(255);
END_VAR
END_METHOD

METHOD ACTIVATEALARM : BOOL
VAR_INPUT
	USIALARMGROUPID : ALARMGROUP_ID;
	UIALARMID : ALARM_ID;
END_VAR
END_METHOD

METHOD ACTIVATEALARMINSTANCE : BOOL
VAR_INPUT
	PFBINSTANCE : POINTER TO BYTE;
	UITEMPLATEALARMID : ALARM_ID;
END_VAR
END_METHOD

METHOD DEACTIVATEALARM : BOOL
VAR_INPUT
	USIALARMGROUPID : ALARMGROUP_ID;
	UIALARMID : ALARM_ID;
END_VAR
END_METHOD

METHOD DEACTIVATEALARMINSTANCE : BOOL
VAR_INPUT
	PFBINSTANCE : POINTER TO BYTE;
	UITEMPLATEALARMID : ALARM_ID;
END_VAR
END_METHOD

METHOD GETALARMIDANDALARMGROUPNAME : BOOL
VAR_INPUT
	UDIALARMGROUPID : UDINT;
	UDIALARMID : UDINT;
END_VAR
VAR_OUTPUT
	SALARMGROUPNAME : STRING;
	UIALARMID : ALARM_ID;
END_VAR
END_METHOD

METHOD GETACTIVEALARMSFROMPROXY
VAR_INPUT
	PASNAME : POINTER TO ARRAY [0..10] OF STRING;
	IGROUPCOUNT : INT;
	FILTERCRITERIA : REFERENCE TO VisuFbAlarmFilterCriteria;
	ITFALARMDATABLOCK : IAlarmDataBlockBaseDINT;
END_VAR
VAR_IN_OUT
	DISTUBPROG : DINT;
END_VAR
END_METHOD

METHOD GETALARMCLASSDESCBYNAMEFROMPROXY
VAR_INPUT
	SPROXYNAME : STRING;
	SCLASSNAME : STRING;
END_VAR
VAR_OUTPUT
	SDESC : ProxyStructAlarmClassDesc;
END_VAR
END_METHOD

METHOD GETALARMCLASSDESCFROMPROXY
VAR_INPUT
	SNAME : STRING;
	UDIID : UDINT;
END_VAR
VAR_OUTPUT
	SDESC : ProxyStructAlarmClassDesc;
END_VAR
END_METHOD

METHOD GETALARMDESCFROMPROXY
VAR_INPUT
	SNAME : STRING;
	UDIALMID : UDINT;
	UDIGRPID : UDINT;
END_VAR
VAR_OUTPUT
	SDESC : ProxyStructAlarmDesc;
END_VAR
END_METHOD

METHOD GETALARMDISPLAYOPTIONSFROMPROXY
VAR_INPUT
	ITFALARMMETAOBJECTSTUB5 : IAlarmMetaObjectStub5;
	REFDISPLAYOPTIONS : REFERENCE TO DisplayOptions;
END_VAR
VAR_OUTPUT
	XVALID : BOOL;
	SCLASSREMAP : STRING;
END_VAR
END_METHOD

METHOD GETALARMGROUPDESCBYNAMEFROMPROXY
VAR_INPUT
	SPROXYNAME : STRING;
	SGRPNAME : STRING;
END_VAR
VAR_OUTPUT
	SDESC : ProxyStructAlarmGroupDesc;
END_VAR
END_METHOD

METHOD GETALARMGROUPDESCFROMPROXY
VAR_INPUT
	SNAME : STRING;
	UDIID : UDINT;
END_VAR
VAR_OUTPUT
	SDESC : ProxyStructAlarmGroupDesc;
END_VAR
END_METHOD

METHOD GETALARMMESSAGEFROMPROXY
VAR_INPUT
	ITFALARMMETAOBJECTSTUB5 : IAlarmMetaObjectStub5;
	IWHICHMESSAGE : INT;
	REFCHARBUFFERSTRING : REFERENCE TO CharBufferString;
	STRINGTYPE : __SYSTEM.TYPE_CLASS;
END_VAR
END_METHOD

METHOD GETALARMMESSAGEFROMPROXY2
VAR_INPUT
	SNAME : STRING;
	STEXTLISTNAME : STRING;
	STEXTLISTINDEX : STRING;
	IWHICHMESSAGE : INT;
	STRINGTYPE : __SYSTEM.TYPE_CLASS;
END_VAR
VAR_OUTPUT
	MESSAGE : CharBufferPtr;
END_VAR
END_METHOD

METHOD GETPROXY : IProxy
VAR_INPUT
	SNAME : STRING;
END_VAR
END_METHOD

METHOD REGISTERALARMCONFIGURATIONREMOTE
VAR_INPUT
	ITFALARMCONFIGURATION : IAlarmConfigurationRemote;
END_VAR
END_METHOD

METHOD SETALARMSTOACKPROXY
VAR_INPUT
	ITFALARMDATABLOCK : IAlarmDataBlockBase2;
END_VAR
END_METHOD

METHOD GETPROXYALARMCLASSESDESCRIPTION : BOOL
VAR_INPUT
	SNAME : STRING;
	PCLDESC : POINTER TO ARRAY [0..0] OF ProxyStructMonitorAlarmClassDesc;
	ISIZE : INT;
END_VAR
VAR_OUTPUT
	ICLCNT : INT;
END_VAR
END_METHOD

METHOD GETPROXYALARMGROUPSDESCRIPTION : BOOL
VAR_INPUT
	SNAME : STRING;
	PGRPDESC : POINTER TO ARRAY [0..0] OF ProxyStructMonitorAlarmGroupDesc;
	ISIZE : INT;
END_VAR
VAR_OUTPUT
	IGRPCNT : INT;
END_VAR
END_METHOD

METHOD GETPROXYALARMSDESCRIPTION : BOOL
VAR_INPUT
	SNAME : STRING;
	PALMDESC : POINTER TO ARRAY [0..0] OF ProxyStructMonitorAlarmDesc;
	DISIZE : DINT;
END_VAR
VAR_OUTPUT
	DIALMCNT : DINT;
END_VAR
END_METHOD

METHOD GETPROXYSTATISTICS : BOOL
VAR_INPUT
	SNAME : STRING;
END_VAR
VAR_OUTPUT
	STRUCTMONITOR : ProxyStructMonitor;
END_VAR
END_METHOD

METHOD GETPROXYSTATISTICSSINGLEACTIVITY : BOOL
VAR_INPUT
	SNAME : STRING;
	ITASKID : INT;
END_VAR
VAR_OUTPUT
	STRUCTMONITOR : ProxyStructMonitorRequest;
END_VAR
END_METHOD

METHOD CLEARTEMPLATEDICTIONARY : BOOL
END_METHOD

METHOD REGISTERTEMPLATEINSTANCE : BOOL
VAR_INPUT
	PINSTANCE : POINTER TO BYTE;
	UDIALARMGROUPID : UDINT;
	UITEMPLATEALARMSOFFSET : UINT;
	UITEMPLATEALARMSLENGTH : UINT;
	PSTALARMTEMPLATENAME : POINTER TO STRING;
	UITEMPLATEEVENTSOFFSET : UINT;
	UITEMPLATEEVENTSLENGTH : UINT;
END_VAR
END_METHOD

METHOD INITAFTERDOWNLOAD : BOOL
END_METHOD

METHOD PRVCHECKALARMMANAGERCLIENT : UDINT
VAR_INPUT
	ITFALARMMANAGERCLIENT : IAlarmManagerClient;
END_VAR
END_METHOD

METHOD PRVCHECKVALIDEVENT : BOOL
VAR_IN_OUT
	UIALARMID : ALARM_ID;
	PALARM8 : IAlarm8;
END_VAR
END_METHOD

METHOD PRVFREECLIENT : UDINT
VAR_INPUT
	PALARMMANAGERCLIENTINFOSTRUCT : POINTER TO AlarmManagerClientInfoStruct;
END_VAR
END_METHOD

METHOD PRVNOTIFYALARMMANAGERCLIENT
VAR_INPUT
	ITFALARMMANAGERCLIENT : IAlarmManagerClient;
	ITFALARM4 : IAlarm4;
END_VAR
END_METHOD

(* ---- STATECOMPARER.fb ---- *)
FUNCTION_BLOCK STATECOMPARER EXTENDS TSLastComparer
END_FUNCTION_BLOCK

METHOD COMPARE : INT
VAR_INPUT
	DIINDEXALARM1 : DINT;
	DIINDEXALARM2 : DINT;
END_VAR
END_METHOD

(* ---- STATISTICS_LTIME.fb ---- *)
FUNCTION_BLOCK STATISTICS_LTIME
VAR_INPUT
	XENABLE : BOOL;
	LTINPUT : LTIME;
END_VAR
VAR
	LTMIN : LTIME;
	LTMAX : LTIME;
	LTAVERAGE : LTIME;
	LICOUNTER : LINT;
	LISUM : LINT;
	XOLDENABLE : BOOL;
	LIAVERAGE : LINT;
	AVERAGE : LTIME;
	COUNT : LINT;
	MAXIMUM : LTIME;
	MINIMUM : LTIME;
END_VAR
END_FUNCTION_BLOCK

(* ---- STRINGCONTAINER.fb ---- *)
FUNCTION_BLOCK STRINGCONTAINER
VAR
	M_BUFFERVECTOR : StringContainerBufferVector;
	M_UDINEXTALLOCATIONSIZE : UDINT := INITIAL_BUFFER_SIZE;
	COMPONENT : STRING := 'StringContainer';
	STRINGTYPE_STRING : UINT := 16;
	STRINGTYPE_WSTRING : UINT := 17;
	INITIAL_BUFFER_SIZE : UDINT := 512;
END_VAR
END_FUNCTION_BLOCK

METHOD ADDSTRING : CharBufferPtr
VAR_INPUT
	CBPMESSAGE : CharBufferPtr;
	TYPECLASS : __SYSTEM.TYPE_CLASS;
END_VAR
VAR_OUTPUT
	UDIERROR : UDINT;
	DISTRINGLENGTH : DINT;
END_VAR
END_METHOD

METHOD FB_EXIT : BOOL
VAR_INPUT
	BINCOPYCODE : BOOL;
END_VAR
END_METHOD

METHOD PRVALLOCATEBUFFER : UDINT
END_METHOD

METHOD PRVALLOCATEBUFFERIFNEEDED : UDINT
END_METHOD

METHOD PRVFINDSTRINGINBUFFER : POINTER TO BYTE
VAR_INPUT
	CBPMESSAGE : CharBufferPtr;
	TYPECLASS : __SYSTEM.TYPE_CLASS;
	UDIWHICHBUFFER : UDINT;
END_VAR
VAR_OUTPUT
	XFOUND : BOOL;
END_VAR
END_METHOD

METHOD PRVHASFREECAPACITY : BOOL
VAR_INPUT
	DICOUNTBYTESREQUIRED : DINT;
	UDIWHICHBUFFER : UDINT;
END_VAR
END_METHOD

METHOD PRVOPENBUFFER : StringContainerBufferInfo
VAR_INPUT
	UDIWHICHBUFFER : UDINT;
END_VAR
END_METHOD

METHOD PRVSTORESTRINGINBUFFER : POINTER TO BYTE
VAR_INPUT
	CBPMESSAGE : CharBufferPtr;
	UISTRINGTYPE : UINT;
	DICOUNTBYTESTOCOPY : DINT;
	DICOUNTBYTESFORSTRING : DINT;
	UDIWHICHBUFFER : UDINT;
END_VAR
END_METHOD

(* ---- STRINGCONTAINERBUFFERVECTOR.fb ---- *)
FUNCTION_BLOCK STRINGCONTAINERBUFFERVECTOR EXTENDS BaseVector
VAR
	_PAPBYSTRINGCONTAINERBUFFERS : POINTER TO ARRAY [0..MAX_NUM_ENTRIES] OF POINTER TO BYTE;
	MAX_NUM_ENTRIES : INT := 10;
END_VAR
END_FUNCTION_BLOCK

METHOD ADDSTRINGCONTAINERBUFFER : UDINT
VAR_INPUT
	PBYBUFFER : POINTER TO BYTE;
END_VAR
END_METHOD

METHOD GETSTRINGCONTAINERBUFFERAT : POINTER TO BYTE
VAR_INPUT
	UDIINDEX : UDINT;
END_VAR
VAR_OUTPUT
	UDIRESULT : UDINT;
END_VAR
END_METHOD

METHOD ABSTRASSIGN : UDINT
VAR_INPUT
	PBT : POINTER TO BYTE;
	UDIINDEX : UDINT;
END_VAR
END_METHOD

METHOD ABSTRDATAPTRCHANGED : UDINT
END_METHOD

METHOD ABSTRSIZEOFELEMENT : UDINT
END_METHOD

(* ---- TEXTHELPER.fb ---- *)
FUNCTION_BLOCK TEXTHELPER
VAR_OUTPUT
	TEXT : STO.TEXT;
END_VAR
END_FUNCTION_BLOCK

METHOD FB_EXIT : BOOL
VAR_INPUT
	BINCOPYCODE : BOOL;
END_VAR
END_METHOD

METHOD FROMSTRING : STO.ERROR
VAR_INPUT
	PS : POINTER TO STRING;
	FUNCTIONCALLER : INT;
END_VAR
END_METHOD

METHOD FROMWSTRING : STO.ERROR
VAR_INPUT
	PWS : POINTER TO WSTRING;
	FUNCTIONCALLER : INT;
END_VAR
END_METHOD

METHOD RELEASE
END_METHOD

(* ---- TIMESTAMPANDVALUESCONTAINER.fb ---- *)
FUNCTION_BLOCK TIMESTAMPANDVALUESCONTAINER
VAR
	M_LITIMESTAMPLAST : AlarmManager_Interfaces.Timestamp;
	M_LITIMESTAMPACTIVE : AlarmManager_Interfaces.Timestamp;
	M_LITIMESTAMPINACTIVE : AlarmManager_Interfaces.Timestamp;
	M_LITIMESTAMPACKNOWLEDGE : AlarmManager_Interfaces.Timestamp;
	M_TRIGGERVALUE : ValueTypeBundle;
	M_ALATCHVARIABLES : ARRAY [1..COUNT_LATCH_VARIABLES] OF ValueTypeBundle;
	COUNT_LATCH_VARIABLES : INT := 10;
END_VAR
END_FUNCTION_BLOCK

METHOD FILL : BOOL
VAR_INPUT
	ITFRANDOMALARMREADACCESS : IRandomAlarmReadAccess;
	DIINDEXALARM : DINT;
	ICOUNTLATCHVARIABLES : INT;
END_VAR
END_METHOD

METHOD GETCOUNTLATCHVARIABLES : USINT
END_METHOD

METHOD GETLATCHVARVALUE : AlarmManagerInternal_Interfaces.ITypedValue2
VAR_INPUT
	IWHICHLATCHVAR : INT;
END_VAR
END_METHOD

METHOD GETCURRENTVALUE : AlarmManagerInternal_Interfaces.ITypedValue
END_METHOD

METHOD GETLATCHVAR1VALUE : AlarmManager_Interfaces.ITypedValue
END_METHOD

METHOD GETLATCHVAR2VALUE : AlarmManager_Interfaces.ITypedValue
END_METHOD

METHOD GETTIMESTAMPACKNOWLEDGE : AlarmManager_Interfaces.Timestamp
END_METHOD

METHOD GETTIMESTAMPACTIVE : AlarmManager_Interfaces.Timestamp
END_METHOD

METHOD GETTIMESTAMPINACTIVE : AlarmManager_Interfaces.Timestamp
END_METHOD

METHOD GETTIMESTAMPLAST : AlarmManager_Interfaces.Timestamp
END_METHOD

METHOD GETTRIGGERVALUE : AlarmManager_Interfaces.ITypedValue
END_METHOD

METHOD GETALARMGROUP : STRING
END_METHOD

METHOD GETCHECKSUM : UDINT
END_METHOD

METHOD GETID : AlarmManager_Interfaces.ALARM_ID
END_METHOD

METHOD GETSTATE : INT
END_METHOD

METHOD SETACKNOWLEDGE
VAR_INPUT
	BACKNOWLEDGEMULTIPLE : BOOL;
END_VAR
END_METHOD

METHOD SETALARMGROUP
VAR_INPUT
	SALARMGROUP : STRING;
END_VAR
END_METHOD

METHOD SETID
VAR_INPUT
	UIID : AlarmManager_Interfaces.ALARM_ID;
END_VAR
END_METHOD

METHOD SETLATCHVAR1VALUE
VAR_INPUT
	ITFTYPEDVALUELATCHVAR1 : AlarmManager_Interfaces.ITypedValue;
END_VAR
END_METHOD

METHOD SETLATCHVAR2VALUE
VAR_INPUT
	ITFTYPEDVALUELATCHVAR2 : AlarmManager_Interfaces.ITypedValue;
END_VAR
END_METHOD

METHOD SETLATCHVARVALUE
VAR_INPUT
	IWHICHLATCHVAR : INT;
	ITFTYPEDVALUELATCHVAR : AlarmManagerInternal_Interfaces.ITypedValue;
END_VAR
END_METHOD

METHOD SETSTATE
VAR_INPUT
	ISTATE : INT;
END_VAR
END_METHOD

METHOD SETTIMESTAMPACKNOWLEDGE
VAR_INPUT
	LITIMESTAMPACKNOWLEDGE : AlarmManager_Interfaces.Timestamp;
END_VAR
END_METHOD

METHOD SETTIMESTAMPACTIVE
VAR_INPUT
	LITIMESTAMPACTIVE : AlarmManager_Interfaces.Timestamp;
END_VAR
END_METHOD

METHOD SETTIMESTAMPINACTIVE
VAR_INPUT
	LITIMESTAMPINACTIVE : AlarmManager_Interfaces.Timestamp;
END_VAR
END_METHOD

METHOD SETTIMESTAMPLAST
VAR_INPUT
	LITIMESTAMPLAST : AlarmManager_Interfaces.Timestamp;
END_VAR
END_METHOD

METHOD SETTRIGGERVALUE
VAR_INPUT
	ITFTYPEDVALUETRIGGER : AlarmManager_Interfaces.ITypedValue;
END_VAR
END_METHOD

(* ---- TL_ALARMSTATUS.fb ---- *)
FUNCTION_BLOCK TL_ALARMSTATUS
VAR
	M_TEXTLISTFILE : STRING(255);
	_STNAMESPACE : STRING;
END_VAR
END_FUNCTION_BLOCK

(* ---- TSACKCOMPARER.fb ---- *)
FUNCTION_BLOCK TSACKCOMPARER EXTENDS AbstractTimestampComparer
END_FUNCTION_BLOCK

METHOD PROTGETTIMESTAMP : BOOL
VAR_INPUT
	DIINDEXALARM : DINT;
END_VAR
VAR_OUTPUT
	LITIMESTAMP : TIMESTAMP;
END_VAR
END_METHOD

(* ---- TSACTIVECOMPARER.fb ---- *)
FUNCTION_BLOCK TSACTIVECOMPARER EXTENDS AbstractTimestampComparer
END_FUNCTION_BLOCK

METHOD PROTGETTIMESTAMP : BOOL
VAR_INPUT
	DIINDEXALARM : DINT;
END_VAR
VAR_OUTPUT
	LITIMESTAMP : TIMESTAMP;
END_VAR
END_METHOD
